        for _i, _step in enumerate(plan, 1):
            _q_raw = list(_step['joints'])
            _q_near = _nearest_in_limit(_q_raw)
            if _q_near != _q_raw:
                log('段%d 关节取同角等价表示：%s → %s'
                    % (_i, ['%.2f' % v for v in _q_raw], ['%.2f' % v for v in _q_near]))
                _step['joints'] = _q_near[:]          # 执行也用归一化值 ✓
            if not _real_limit_ok(_step['joints'], _lo, _hi):
                raise ValueError('段%d 目标关节超出实机限位：%s（规划期应已过滤，此为最后防线；已试 ±360 同角表示）'
                                 % (_i, ['%.2f' % v for v in _step['joints']]))
        for before, after in ((frame, robot.PoseFrame()), (tool, robot.PoseTool())):
            error = invH(before)*after
            if norm(error.Pos()) > 0.01 or pose_angle(error) > math.radians(0.01):
                raise RuntimeError('预检期间工具或参考坐标系改变，取消执行。')
        robot.setSpeed(ROBOT_SPEED)
        RDK.Command('Trace','Reset')
        RDK.Command('Trace','On')
        expected = start
        # v14k：停用长运动分瓣（split_moves 恒 False）。2026-10-12 实测日志坐实：假断连与跨度无关，
        # 60°/95°/169°/180° 的瓣与 20mm 途经点每条指令都在断，分瓣已不防任何东西，只剩每瓣一轮
        # 等待+重连停顿税；_single_move_settle 断连容忍（_wait_controller_static 20s 静止上限）
        # 罩得住单条长指令的收尾（20°/s 下 180°≈9s<20s）。分瓣机制与常量原样留档，遇真断连指纹
        # （未自然收尾/未到位）随时把本行改回 single_method is None and len(records) > 1 即可恢复。
        split_moves = False
        movl_direct = bool(real_movldirect_var.get()) if _movl_direct_ready() else False
        if movl_direct:
            # v15：原来的超长版本横幅已按用户要求删除，只留一行关键参数，便于判读
            log('直发开启 ｜ 段长≤%.0fmm ｜ 法兰容差 %.0fmm/%.1f° ｜ 等待≤%.0fs ｜ 禁直发名单=%s'
                % (MOVL_DIRECT_MAX_MM, MOVL_FLANGE_TOL_MM, MOVL_FLANGE_TOL_DEG,
                   MOVL_ARRIVE_WAIT_S, MOVL_DIRECT_BLOCK_POINTS))
        log('本次单条MovL动态认证放行点=%s' % [i for i,s in enumerate(plan,1) if s.get('direct_movl_certified')])
        _assert_continuous_dispatch(records, start, plan, movl_direct)
        for i, step in enumerate(plan, 1):
            for rewind in step['rewinds']:
                _require_joints(expected)
                _move_with_completion_check("MoveJ", rewind, split_moves)
                _require_joints(rewind)
                expected = rewind
            _require_joints(expected)
            waypoints = step.get('waypoints') or []
            if step['method'] == 'MoveL' and not waypoints:
                # 理论不可达：v13 起所有 MoveL 步都带细分途经点；不带则说明规划层契约被破坏
                raise RuntimeError(f"P{i}：MoveL 步缺少细分途经点，拒绝发送驱动 MOVL（已判死）。")
            seg_mm = seg_rot = None
            if movl_direct and step['method'] == 'MoveL' and waypoints:
                # 仅开关开启时才算（两次 FK 的 API 往返）；开关关/离线 verify 零开销
                _seg_rel = _trajectory_pose(step['joints']) * invH(_trajectory_pose(expected))
                seg_mm, seg_rot = norm(_seg_rel.Pos()), pose_angle(_seg_rel)
            direct_ready = (movl_direct and _direct_step_allowed(i, step)
                            and seg_mm is not None
                            and seg_mm <= MOVL_DIRECT_MAX_MM
                            and seg_rot <= math.radians(0.5))
            _send_q = step.get('direct_send_joints', step['joints'])
            if direct_ready and not step.get('direct_movl_certified'):
                # v14w：发送前数字净化——控制器 -30001 拒的是【参数形态】不是几何（LOG_VERSION
                # 处 11:38 拒收 / 15:55 接受两份实录）。净化只在零边界区微调发送关节；
                # 净化失败 ⇒ direct_ready=False ⇒ 落到 elif waypoints 走细分（安全回落）。
                _send_q, _purge_note = _movl_digit_safe_joints(step['joints'])
                if _send_q is None:
                    log('P%d：⛔ %s ⇒ 改走细分途经点路径。' % (i, _purge_note))
                    direct_ready = False
                elif _purge_note:
                    log('P%d：%s' % (i, _purge_note))
            if direct_ready:
                # v14p 法兰补偿MOVL：驱动 MOVL 无工具补偿、按法兰执行（v14l 11:30 实证停点法兰=
                # 命令TCP目标，差仅5.5mm）——将错就错：把本步构型的【法兰位姿】直接当笛卡尔目标
                # 发给控制器，法兰被精确送到位，物理工具尖端（182mm，v14w27 实测）随之落在认证
                # 直线上。姿态恒定段法兰线=TCP线平移常向量，扫掠包络与细分路径一致。
                # v14w36/37 演进：v14w36 只改传位姿（不切工具）⇒ MoveL(位姿) 按 TCP 空间
                # 校验，P8 法兰位姿被反推到 z=744 爆臂展 TargetReachError（11:18 实录）；
                # v14w37 = 位姿传递（动画=认证直线，根治关节弧假碰撞冻死）+ 发送窗口单位
                # 变换（校验/数字=法兰空间）；柜子实收参数与旧金标准逐位一致（0 偏差）。
                log(f"P{i}：v14w 法兰补偿MOVL：段长{seg_mm:.1f}mm（姿态变化{math.degrees(seg_rot):.2f}°），收起 {len(waypoints)} 个细分途经点，一指令直发（发法兰位姿=自算FK+单位变换窗口，发送关节已净化；v14w37）。")
                # v14r：require_joints=False——假断连分支的关节级 0.5° 校验让位给下方
                # 法兰级粗验收+MoveJ 微纠偏收口（终点仍回认证构型，护栏语义不降级）。
                # v14u：expect_target=段目标关节——目标锚定到位等待（上限 60s，每5s进度日志）。
                # v14w：净化只作用于发送关节；expect_target 仍是认证关节（到位判据不变）。
                # v14w37：位姿传递（动画=认证直线）+ flange_space 单位变换（校验/数字=法兰空间）。
                _send_pose = invH(robot.PoseFrame()) * robot.SolveFK(_send_q)
                # ★ 2026-11-03（可选，默认关）：先给控制器发 Tool(0)/User(0)，
                # 治 `[MovL#878] movL not set tool or user!!!` ⇒ 让 MovL 明确按 基座系+零工具(法兰) 执行。
                # 打开方式：把 MOVL_SEND_TOOL_USER 改成 True（建议先跑一条短段验证）。
                if MOVL_SEND_TOOL_USER:
                    if _try_set_tool_user():
                        log('  ✓ Tool(0)/User(0) 已下发，继续直发')
                    else:
                        raise ControllerMotionFault('Tool/User未确认，停止直发。')
                log('P%d：发送法兰目标=%s；认证关节=%s；TCP=%s' % (i, Pose_2_Fanuc(_send_pose), step['joints'], Pose_2_Fanuc(robot.PoseTool())))
                _single_move_settle('MoveL', _send_pose, require_joints=False,
                                    expect_target=step['joints'], flange_space=True)
                # ★★★ v15.7（2026-11-03）：直发结束后【先等真静止】再做后续（法兰验收/收口）。
                #   实录（v15.6, P8）：直发报"已完成"（假断连分支）→ 脚本立刻法兰验收(5.71mm ✓)
                #   → P8 尾部关节检查【通过】（读到的是过渡中姿态）→ P9 开头再读【已翻转】⇒ 差 20~38° ⇒ 停 ✗
                #   对比：P7 目标 [75.42,12.24,57.74,20.02] vs 停止实测 [78.10,36.86,19.48,33.66]
                #         ⇒ J2↑25 / J3↓38 / J4↑14 = 典型【肘部翻转 elbow flip】✗
                #   机理：MovL 只给位姿 ⇒ 控制器自行选 IK 分支（可能选翻转那组）✗
                #         + 直发"已完成"没等真静止 ⇒ 后续读到的是过渡值 ✗
                #   ⇒ 这里补一段【关节稳定等待】：连续 3 次采样（每次 0.3s）关节变化 <0.05° 才算真停，
                #     最多等 8 秒；等稳定后再做验收/收口，避免"读到过渡值"造成的假通过/假失败。
                _st = None
                _stable = False
                for _w in range(24):          # 24 × 0.3s ≈ 7.2s 上限
                    _cur = _live_joints()
                    if _st is not None and max(abs(a - b) for a, b in zip(_cur, _st)) < 0.05:
                        _stable = True
                        break
                    _st = _cur
                    time.sleep(0.3)
                if not _stable:
                    log('P%d：⚠️ 直发后 7 秒内关节仍未稳定（继续按现值验收，可能判死）' % i)
                else:
                    log('P%d：直发后关节已稳定 ✓（进入法兰验收/收口）' % i)
                # ★★★ v15.8（2026-11-03）：★ 安全网 —— 直发是【控制器自行选 IK 解】，
                #   规划期的自干涉硬禁区（|J4|>150 等）拦不到它 ✗
                #   ⇒ 直发落点若真落进禁区（J4 极端 / J4×J5 组合区），必须【立刻回认证构型】，
                #     绝不能把手臂留在危险姿态里继续跑下一段 ✓
                _post = _live_joints()
                if _real_interfere_combo(_post):
                    log('P%d：🚨 直发落点落入自干涉禁区！实测=%s（J4=%.2f J5=%.2f）⇒ 立即回认证构型'
                        % (i, ['%.2f' % v for v in _post], _post[3], _post[4]))
                    _single_move_settle('MoveJ', step['joints'])
                    _require_joints(step['joints'])
                    log('P%d：已回到认证构型 ✓' % i)
                elif abs(_post[3]) > REAL_INTERFERE_J4_MAX:
                    log('P%d：⚠️ 直发落点 J4=%.2f° 偏大（>%.0f° 组合区阈值，但未触禁区组合）——记录'
                        % (i, _post[3], REAL_INTERFERE_J4_MAX))
                try:
                    robot.setJoints(_post)   # 显示实测姿态，不用预期目标掩盖未到位。
                except Exception:
                    pass
                # v14q：MovL 落点法兰级粗验收（≤8mm/≤1°）+ MoveJ 微纠偏收口（关节级 0.5° 罩终点）。
                # v14p 首航停在 0.95° 关节残差（法兰 4.61mm/0.616°）被 0.5° 护栏拦停——那是控制器
                # MovL 固有落点残差（v14l 5.5mm 双样本背书），不是构型错误；但终点必须回到认证构型，
                # 故验收通过后用一条短 MoveJ（~1° 关节差）收口，走 _single_move_settle 全套护栏。
                _actual, _is_static = _wait_controller_static(samples=3, interval=0.2)
                _mm, _deg = _movl_flange_accept(_actual, step['joints'])
                if _mm > MOVL_FLANGE_TOL_MM or _deg > MOVL_FLANGE_TOL_DEG:
                    raise RuntimeError('v14u 法兰级粗验收未过：停点法兰残差%.2fmm/%.2f°（容差%.1fmm/%.1f°），实测关节%s，停止待判读。'
                                       % (_mm, _deg, MOVL_FLANGE_TOL_MM, MOVL_FLANGE_TOL_DEG,
                                          ['%.2f' % v for v in _actual]))
                _jm = max(abs(a - b) for a, b in zip(_actual, step['joints']))
                if _jm > MOVE_OFFSET_TOL:
                    log(f"P{i}：v14u MovL 直发落点法兰级验收通过（残差{_mm:.2f}mm/{_deg:.2f}°），关节残差{_jm:.2f}°——发 MoveJ 微纠偏收口。")
                    # ★★★ v15.4（2026-11-03）：收口 MoveJ 加重试 —— 治"P8 停下"：
                    #   实录 11:29:03 验收通过 → 发收口 MoveJ → 11:29:04 驱动报断连 → 11:29:06 才重连
                    #   ⇒ 那条收口 MoveJ 没走完 ⇒ 关节残差 2.68° 残留
                    #   ⇒ 下一段前的 _require_joints（容差 0.5°）判死 ⇒ 停在 P8 ✗
                    #   收口目标是【认证构型】（确定可达）⇒ 重发安全 ✓；最多 2 次，仍不到就抛原错。
                    _close_err = None
                    for _close_try in (1, 2):
                        try:
                            _single_move_settle('MoveJ', step['joints'])
                            _close_err = None
                            break
                        except Exception as _close_exc:  # noqa: BLE001
                            _close_err = _close_exc
                            if _close_try == 1:
                                log('P%d：收口 MoveJ 未完成（%s: %s）⇒ 重试一次（目标为认证构型，可达）'
                                    % (i, type(_close_exc).__name__, _close_exc))
                                time.sleep(0.5)
                    if _close_err is not None:
                        raise _close_err
                # ★★★ v15.5（2026-11-03）：直发+收口之后，再做【关节校正重试】—— 治 P8 停下的真因。
                #   实录（v15.4, 11:36:19~23）：
                #     P8 直发到位（关节残差 2.68°）→ 法兰验收通过 → 发收口 MoveJ
                #     → 驱动报断连 → 脚本打印「驱动断连但运动已自然完成到位」（★ 它认为完成 ✗）
                #     → 于是 _single_move_settle 没抛异常（断连分支 require_joints=False 不校验关节）
                #     → 紧接的 _require_joints 才发现不一致（实测 J2=36.86/J3=19.48，差很多）⇒ 抛错停 ✗
                #   ⇒ 所以 v15.4 的 try/except 重试【根本没触发】✗
                #   ⇒ 改为：_require_joints 失败时【再发一次定向 MoveJ】校正（目标=认证构型，确定可达）
                try:
                    _require_joints(step['joints'])
                except Exception:
                    log('P%d：直发+收口后关节仍与预检不一致 ⇒ 再发一次 MoveJ 校正（目标为认证构型，可达）' % i)
                    time.sleep(0.5)
                    _single_move_settle('MoveJ', step['joints'])
                    _require_joints(step['joints'])
                    log('P%d：校正 MoveJ 完成 ✓' % i)
            elif (movl_direct and not _direct_step_allowed(i, step) and seg_mm is not None
                    and seg_mm <= MOVL_DIRECT_MAX_MM and seg_rot <= math.radians(0.5)):
                # ★ v14v4：本点被【禁直发名单】拦下 —— 明确告知，便于判读日志
                log(f"P{i}：⛔ 本点在【禁直发名单】MOVL_DIRECT_BLOCK_POINTS={MOVL_DIRECT_BLOCK_POINTS} 里 ⇒ "
                    f"不走法兰补偿直发，改走【细分途经点路径】（v14n 实测 17/17 通过、零事故的路径）。")
                if not waypoints:
                    raise RuntimeError(f'P{i}：禁直发点缺少途经点，停止。')
                for way in waypoints:
                    _move_with_completion_check('MoveJ', way, False)
                    _require_joints(way)
                _require_joints(step['joints'])
            elif waypoints:
                log(f"P{i}：执行预检方案 {step['method']}→MoveJ 细分，{len(waypoints)} 个途经点，终点关节={step['joints']}")
                for k, way in enumerate(waypoints, 1):
                    _move_with_completion_check('MoveJ', way, False)
                    _require_joints(way)
                _require_joints(step['joints'])
            else:
                log(f"P{i}：执行预检方案 {step['method']}，关节={step['joints']}")
                _move_with_completion_check(step['method'], step['joints'], split_moves)
                _require_joints(step['joints'])
            expected = step['joints']
            completed += 1
        log(f'实机执行完成：{completed}/{len(plan)}点。')
    except Exception as exc:
        log(f'实机任务停止，已完成{completed}点：{type(exc).__name__}: {exc}')
        if movl_direct and ('断连' in str(exc) or '未到位' in str(exc) or '落点偏差' in str(exc) or '粗验收' in str(exc)):
            log('【v14u】法兰补偿MOVL执行段出断连/落点指纹（v14w24 无勾选框；细分途经点路径保留在计划中，可作回退依据）。')
        try:
            actual, velocity, mode = _controller_feedback()
            log('停止时控制器实际反馈：关节=%s，速度=%s，模式=%s；不自动重发运动。' % (actual, velocity, mode))
        except Exception as feedback_error:
            log('停止时也无法取得控制器反馈：%s' % feedback_error)
    finally:
        _real_running = False
        try:
            _keepalive_stop.set()
            _ka_thread.join(timeout=3)
        except Exception:
            pass


def _point_to_segment_distance(p, a, b):
    """3D点到线段距离，单位mm。"""
    ax, ay, az = a
    bx, by, bz = b
    px, py, pz = p
    ab = (bx-ax, by-ay, bz-az)
    ap = (px-ax, py-ay, pz-az)
    ab2 = ab[0]*ab[0] + ab[1]*ab[1] + ab[2]*ab[2]
    if ab2 < 1e-12:
        return math.sqrt((px-ax)**2 + (py-ay)**2 + (pz-az)**2)
    t = (ap[0]*ab[0] + ap[1]*ab[1] + ap[2]*ab[2]) / ab2
    t = max(0.0, min(1.0, t))
    q = (ax+t*ab[0], ay+t*ab[1], az+t*ab[2])
    return math.sqrt((px-q[0])**2 + (py-q[1])**2 + (pz-q[2])**2)


def _tcp_position_from_joints(q):
    """关节角 -> 当前参考坐标系下的TCP位置，与轨迹输入使用同一坐标系。"""
    f = pose_to_fanuc_values(invH(robot.PoseFrame()) * robot.SolveFK(q) * robot.PoseTool())
    return (float(f[0]), float(f[1]), float(f[2]))


def _check_movej_tcp_trajectory(start_q, target_q, start_tcp_vals, target_tcp_vals, log, samples=30, max_deviation_mm=None):
    """
    在真正执行MoveJ之前，用关节空间线性插补采样，计算TCP轨迹相对
    起点-终点TCP直线段的最大偏离距离。

    目的：MoveL失败时，不再无条件MoveJ；只有MoveJ造成的TCP空间绕行
    没有超过允许值，才允许用MoveJ兜底。
    """
    if max_deviation_mm is None:
        max_deviation_mm = MOVEJ_FALLBACK_MAX_DEVIATION_MM

    start_q = [float(v) for v in start_q[:6]]
    target_q = [float(v) for v in target_q[:6]]
    a = (float(start_tcp_vals[0]), float(start_tcp_vals[1]), float(start_tcp_vals[2]))
    b = (float(target_tcp_vals[0]), float(target_tcp_vals[1]), float(target_tcp_vals[2]))

    log("开始检查 MoveJ 兜底轨迹：%d 个采样点，允许最大TCP偏离 %.3f mm" % (samples + 1, max_deviation_mm))
    max_dev = -1.0
    max_info = None

    for k in range(samples + 1):
        t = float(k) / float(samples)
        q = [start_q[j] + (target_q[j] - start_q[j]) * t for j in range(6)]
        try:
            p = _tcp_position_from_joints(q)
        except Exception as e:
            log("  MoveJ轨迹检查失败：第 %d/%d 个采样点 FK失败：%s: %s" % (k+1, samples+1, type(e).__name__, e))
            return False

        dev = _point_to_segment_distance(p, a, b)
        if dev > max_dev:
            max_dev = dev
            max_info = (k, t, q, p)

        if dev > max_deviation_mm:
            log("✕ MoveJ兜底轨迹拒绝：第 %d/%d 个采样点偏离TCP直线 %.3f mm > %.3f mm" %
                (k+1, samples+1, dev, max_deviation_mm))
            log("  t=%.3f  TCP=(%.3f, %.3f, %.3f)" % (t, p[0], p[1], p[2]))
            log("  因此不会执行这个MoveJ兜底动作，避免出现不可接受的大绕圈。")
            return False

    if max_info is not None:
        k, t, q, p = max_info
        log("✓ MoveJ兜底轨迹检查通过")
        log("  最大TCP偏离直线：%.3f mm（采样 %d/%d，t=%.3f）" % (max_dev, k+1, samples+1, t))
        log("  最大偏离点TCP=(%.3f, %.3f, %.3f)" % (p[0], p[1], p[2]))
    return True


# ============================================================
# 执行连续运动（MoveL失败时先检查MoveJ轨迹）
# ============================================================
def _collision_details():
    pairs = RDK.CollisionPairs()
    return '；'.join(f'{a.Name()}[连杆{ia}] 与 {b.Name()}[连杆{ib}]'
                    for a, b, ia, ib in pairs) or '路径碰撞或关节不可行'


def _enable_obstacle_checks():
    if RDK.RunMode() != RUNMODE_SIMULATE:
        raise RuntimeError('障碍物预检仅允许在仿真模式执行。')
    # 每次进入预检都清空预检缓存：缓存生命周期 = 单次预检规划，
    # 障碍物/工作站状态的变化在下一次预检即时生效。
    _plan_cache.clear()
    for name in ('安装台_650x650x80mm', '地面_禁止穿越', '磨砂圆柱_R150_H50', '挡板_半封闭3面'):
        obstacle = RDK.Item(name, ITEM_TYPE_OBJECT)
        if not obstacle.Valid():
            raise RuntimeError(f'缺少障碍物模型：{name}，请加载包含台子和地面的工作站。')
        if name == '安装台_650x650x80mm':
            if RDK.setCollisionActivePair(COLLISION_OFF, robot, obstacle, 0, 0) != 1:
                raise RuntimeError('无法配置安装台与固定底座的接触关系。')
        for link in range(1, 7):
            if RDK.setCollisionActivePair(COLLISION_ON, robot, obstacle, link, 0) != 1:
                raise RuntimeError(f'无法启用{name}与连杆{link}的碰撞检查。')
        tool_items = list(RDK.ItemList(ITEM_TYPE_TOOL))
        _handle = RDK.Item('门把手_bs1')   # v14w12：网格替换后可能为 OBJECT 类型，按名并入
        if _handle.Valid() and all(_handle.item != t.item for t in tool_items):
            tool_items.append(_handle)
        for tool in tool_items:
            parent = tool.Parent()
            while parent.Valid() and parent.item != robot.item:
                parent = parent.Parent()
            if parent.Valid() and RDK.setCollisionActivePair(COLLISION_ON, tool, obstacle) != 1:
                raise RuntimeError(f'无法启用{name}与工具的碰撞检查。')
    RDK.setCollisionActive(COLLISION_ON)


def _check_single_joint_path(end):
    _enable_obstacle_checks()
    saved = robot.Joints().list()[:6]
    try:
        RDK.Command('Trace', 'Off')
        RDK.Render(False)
        if _movej_test_cached(saved, end, 1) != 0:
            raise ValueError('单点MoveJ路径被拒绝：' + _collision_details())
    finally:
        robot.setJoints(saved)
        RDK.Render(True)


def _trajectory_pose(q):
    return invH(robot.PoseFrame()) * robot.SolveFK(q) * robot.PoseTool()


def _reorient_next_pose(records, i, rec):
    """v14w33：i 为 1-based 点号。若下一点存在且为【同 TCP 位姿纯换姿】（xyz 全同、姿态不同），
    返回下一点的 TCP 位姿 Mat，否则 None。用于换姿对的分支前视。"""
    try:
        if i >= len(records):
            return None
        nxt = records[i]          # 0-based 列表：下一条记录
        if nxt['type'] != 'TCP' or nxt.get('singular', False):
            return None
        va = [float(v) for v in rec['values'][:6]]
        vb = [float(v) for v in nxt['values'][:6]]
        if all(abs(va[k] - vb[k]) < 1e-9 for k in range(3)) and any(abs(va[k] - vb[k]) > 1e-9 for k in range(3, 6)):
            return fanuc_values_to_pose(*vb)
    except Exception:
        return None
    return None


def _linear_path_endpoint(start, target):
    """带结果缓存：分支重试时同一（起点, 目标）不重复计算。"""
    key = ('linear', _cache_key_joints(start), _cache_key_pose(target))
    if key in _plan_cache:
        return _plan_cache[key]
    result = _linear_path_endpoint_uncached(start, target)
    _plan_cache[key] = result
    return result


def _linear_path_endpoint_uncached(start, target):
    # 粗筛：10mm 采样点是 1mm 采样点的子集，粗筛失败则 1mm 细查必然失败，
    # 可直接拒绝；粗筛通过后再跑原有 1mm 细查，通过/拒绝判定与只跑 1mm 完全一致。
    if RDK.RunMode() != RUNMODE_SIMULATE:
        raise RuntimeError('直线路径预检仅允许在仿真模式执行。')
    # v15.17: Lookahead may leave the model at the P10 wrist-spin posture.
    # RoboDK's numerical IK uses current model joints even with an explicit j1.
    # Reset the model seed before each independent path check.
    robot.setJoints(start)
    status = robot.MoveL_Test(start, target, minstep_mm=10)
    if status == 0:
        robot.setJoints(start)
        status = robot.MoveL_Test(start, target, minstep_mm=1)
    if status != 0:
        return None, f'MoveL原生路径检查未通过（{status}）：' + _collision_details()
    # 本机MoveL_Test返回成功后Joints()可能为全零；从插补矩阵读取实际终点。
    # 碰撞判定已由上方同路径 1mm MoveL_Test 完成，此处仅提取终点关节，
    # 关闭碰撞检查提速（实测约快两个数量级）；整段权威碰撞复核仍在
    # _verify_obstacle_plan（碰撞开、1mm）进行。
    program = RDK.AddProgram('_TCP仿真_路径预检', robot)
    try:
        program.setVisible(False)
        robot.setJoints(start)
        program.setPoseFrame(robot.PoseFrame())
        program.setPoseTool(robot.PoseTool())
        program.MoveJ(start)
        program.MoveL(target)
        message, matrix, status = program.InstructionListJoints(mm_step=1, deg_step=1, collision_check=COLLISION_OFF)
        if status < 0:
            return None, message
        end = matrix.tr().rows[-1][:6]
        error_pose = invH(target) * _trajectory_pose(end)
        if norm(error_pose.Pos()) > .01 or pose_angle(error_pose) > math.radians(.01):
            raise RuntimeError('路径预检返回的终点不匹配目标TCP。')
        return end, message
    finally:
        program.Delete()


def _linear_waypoints(start, target, step_mm=None):
    """v13：从一条 MoveL 指令采样细分途经关节点（按 IK 顺序，无分支翻转）。

    用 InstructionListJoints(mm_step=LINEAR_SUBSTEP_MM, collision_check=COLLISION_OFF) 采样：
    途经点与 MoveL 执行的是同一条几何直线，且 IK 连续选解（避免用全局 SolveIK 时
    途经点在多解间跳变）。碰撞已由 _linear_path_endpoint 的 MoveL_Test@1mm 权威判定，
    此处不再重复。返回含终点的关节点列表；空列表表示采样失败（调用方回退直达）。"""
    if step_mm is None:
        step_mm = LINEAR_SUBSTEP_MM
    key = ('waypoints', _cache_key_joints(start), _cache_key_pose(target), round(float(step_mm), 3))
    if key in _plan_cache:
        return [q[:] for q in _plan_cache[key]]
    program = RDK.AddProgram('_TCP仿真_细分采样', robot)
    saved = robot.Joints().list()[:6]
    try:
        program.setVisible(False)
        robot.setJoints(start)
        program.setPoseFrame(robot.PoseFrame())
        program.setPoseTool(robot.PoseTool())
        program.MoveJ(start)
        program.MoveL(target)
        message, matrix, status = program.InstructionListJoints(mm_step=step_mm, deg_step=1, collision_check=COLLISION_OFF)
        cols = matrix.tr().rows if matrix is not None else []
        if status < 0 or not cols:
            return []
        # 丢弃比步长更密的重复点（InstructionListJoints 在奇异附近会加密采样）
        picked = [list(map(float, cols[0][:6]))]
        for row in cols[1:]:
            q = list(map(float, row[:6]))
            if max(abs(a - b) for a, b in zip(q, picked[-1])) >= step_mm / 10.0:
                picked.append(q)
        # 去尾：InstructionListJoints 可能带比目标多一点的收尾点，以关节距离最近的为准
        end_q, _ = _linear_path_endpoint(start, target)
        if end_q is not None and picked and max(abs(a - b) for a, b in zip(end_q, picked[-1])) > 1.0:
            picked[-1] = list(map(float, end_q))
        _plan_cache[key] = [q[:] for q in picked]
        return [q[:] for q in picked]
    finally:
        program.Delete()
        robot.setJoints(saved)


def _obstacle_posture_key(q, reference=None):
    table = RDK.Item('安装台_650x650x80mm', ITEM_TYPE_OBJECT)
    height = 0.0
    if table.Valid():
        elbow = invH(table.PoseAbs()) * robot.PoseAbs() * robot.JointPoses(q)[3]
        height = elbow.Pos()[2]
    return (-round(height, 6), sum((v-r)**2 for v, r in zip(q, reference or [0]*6)), tuple(q))


def _obstacle_joint_target(start, values, max_deviation=None, log=None):
    """带结果缓存：同一（起点, 目标, 偏离上限）的兜底选解不重复搜索。"""
    key = ('obstacle', _cache_key_joints(start), tuple(round(float(v), 6) for v in values[:6]),
           round(float(max_deviation), 6) if max_deviation is not None else None)
    if key in _plan_cache:
        cached = _plan_cache[key]
        if isinstance(cached, ValueError):
            raise cached
        return cached
    try:
        result = _obstacle_joint_target_uncached(start, values, max_deviation, log)
    except ValueError as exc:
        _plan_cache[key] = exc
        raise
    _plan_cache[key] = result
    return result


def _obstacle_joint_target_uncached(start, values, max_deviation=None, log=None):
    # v14-P2P：不再用 seed 候选/肘高排序，直接取离当前关节最近的逆解做逐级检查；
    # 最近解过不了偏离/碰撞时仍会在这里报错（单点 MoveJ 兜底路径保持可用）。
    lower, upper, _ = robot.JointLimits()
    candidates = [_nearest_ik_from_current(start, fanuc_to_pose(*values))]
    saved = robot.Joints().list()[:6]
    try:
        # 少量FK采样仅用于排序；不能替代后面的偏离复核与精细碰撞检查。
        a = _tcp_position_from_joints(start)
        table = RDK.Item('安装台_650x650x80mm', ITEM_TYPE_OBJECT)
        base_to_table = invH(table.PoseAbs()) * robot.PoseAbs()
        ranked = []
        for end in candidates:
            deviation, height = 0.0, float('inf')
            for k in range(11):
                q = [x + (y-x)*k/10 for x, y in zip(start, end)]
                deviation = max(deviation, _point_to_segment_distance(
                    _tcp_position_from_joints(q), a, values[:3]))
                height = min(height, (base_to_table * robot.JointPoses(q)[3]).Pos()[2])
            if max_deviation is not None and deviation > max_deviation:
                continue
            # 20mm一档，避免为很小的偏离差反复搜索；同档优先抬高肘部。
            ranked.append(((int(deviation/20), -height,
                            sum(abs(y-x) for x, y in zip(start, end))), end))
        checked = 0
        for _, end in sorted(ranked, key=lambda entry: entry[0]):
            if max_deviation is not None and not _check_movej_tcp_trajectory(
                    start, end, pose_to_fanuc_values(_trajectory_pose(start)), values,
                    lambda msg: None, samples=100, max_deviation_mm=max_deviation):
                continue
            checked += 1
            if _movej_test_cached(start, end, .25) == 0:
                if log is not None:
                    log(f'MoveJ快速筛选：{len(candidates)}个候选，{len(ranked)}个通过粗筛，精查{checked}条后找到合格路径。')
                return end
        raise ValueError('所有候选关节路径均碰撞、超出偏离限制或没有有效逆解。')
    finally:
        robot.setJoints(saved)


def _verify_obstacle_plan(start, plan):
    program = RDK.AddProgram('_TCP仿真_整段碰撞复核', robot)
    saved = robot.Joints().list()[:6]
    try:
        program.setVisible(False)
        program.setPoseFrame(robot.PoseFrame())
        program.setPoseTool(robot.PoseTool())
        program.MoveJ(start)
        for step in plan:
            for q in step['rewinds']:
                program.MoveJ(q)
            if step['method'] == 'MoveL' and not step.get('waypoints'):
                # v13 防呆：MoveL 步必须带细分途经点，否则规划层契约被破坏
                raise ValueError('整段碰撞复核：MoveL 步缺少细分途经点，拒绝。')
            getattr(program, step['method'])(step['joints'])
        message, matrix, status = program.InstructionListJoints(
            mm_step=1, deg_step=1, collision_check=COLLISION_ON)
        if status < 0 or 'collision' in message.lower():
            raise ValueError('整段碰撞复核未通过：' + message)
    finally:
        program.Delete()
        robot.setJoints(saved)


# Continuous TCP paths always recover calibrated-body IK branches and re-certify
# their actual command paths. Record hashes bind receipts, never enable policy.
CALIBRATED_IK_SEEDS = [[163.62039271007563, 64.01735255223417, -67.25050650734438, 93.2331539551102, -90.00000000000001, -106.37960728992437], [-72.40715810734315, -20.66480267505412, -103.89758096136477, 124.56238363641887, 72.40715810734312, 0.0], [-58.553344176794326, -22.475689666466394, -101.12528805253322, 123.60097771899962, 58.55334417679429, -1.0294949594003553e-14], [-58.553344176794326, -22.475689666466394, -101.12528805253322, 123.60097771899962, 58.55334417679429, 180.0], [-87.40476475829131, -22.47568966646641, -101.12528805253322, 123.60097771899962, 87.40476475829125, 180.0], [-64.66430037296594, -3.2481937678895747, -126.71804809984242, 129.96624186773198, 64.66430037296595, 180.0], [-75.41679324948196, -12.462263518678185, -56.77419042193441, -20.76354605938741, 90.0, 194.58320675051806], [-78.10373775148642, -37.83824919659381, -16.865010237740023, -35.296740565666134, 90.0, 191.89626224851355], [-88.23587605840977, -43.75520866199254, -5.060724146438354, -41.184067191569056, 90.0, 181.7641239415902], [-88.23587605840977, -43.75520866199254, -5.060724146438354, -41.184067191569056, 90.0, 1.7641239415902135], [-68.33462268250656, -43.75520866199333, -5.060724146436616, -41.184067191570016, 89.99999999999999, 21.665377317493437], [61.81374704354286, 48.51918849734889, 55.392423259627606, -103.91161175697648, 28.186252956457167, 180.0], [62.25330564679723, 54.06615976151417, 44.56648765802543, -98.6326474195396, 27.746694353202802, 180.0], [61.81374704354286, 48.51918849734889, 55.392423259627606, -103.91161175697648, 28.186252956457167, 90.0], [62.253305646797244, 54.06615976151415, 44.56648765802541, -98.63264741953954, 27.746694353202788, 89.99999999999999], [61.81374704354286, 48.51918849734889, 55.392423259627606, -103.91161175697648, 28.18625295645714, -90.00000000000001], [62.25330564679723, 54.0661597615141, 44.56648765802556, -98.63264741953965, 27.746694353202773, -90.00000000000004], [62.57433490659918, 47.78974891048301, 57.14855554302247, -103.76676871515006, 27.416346223420135, -60.70732349501101], [62.98154845233014, 53.155168153175346, 46.7150047327387, -98.68233310181975, 27.009218983764953, -60.72565665513798], [62.57582549469282, 48.080389017894106, 56.23528280269005, -104.31567182058413, 27.424174505307207, -180.0], [62.71034615480792, 51.83128832842894, 49.315963732196764, -99.89133677590429, 25.437207443150072, -301.4668568689523], [60.218467190004304, 39.42913510297621, 54.58098026787218, -92.8583848548389, 27.92853761288419, -301.35028218541504], [-13.591622773947876, 18.9460252211274, 48.02925373146127, 23.02472104741136, -90.0, -193.59162277394785]]
_continuous_profile_active = False


def _records_fingerprint(records):
    import hashlib
    canonical = [dict(type=r['type'], values=[0.0 if abs(float(v)) < 1e-12 else float(v)
                 for v in r['values']], singular=bool(r.get('singular', False)),
                 spin360=bool(r.get('spin360', False)), j6_delta=int(r.get('j6_delta', 0)))
                 for r in records]
    return hashlib.sha256(json.dumps(canonical, sort_keys=True,
        separators=(',', ':')).encode('utf-8')).hexdigest()


def _continuous_records(records):
    return len(records) > 1 and any(r.get('type') == 'TCP' for r in records)


def _assert_continuous_dispatch(records, initial, plan, direct_enabled):
    if not _continuous_records(records):
        return
    fingerprint = _records_fingerprint(records)
    previous = initial
    for number, step in enumerate(plan, 1):
        if step.get('waypoints'):
            certificate = step.get('direct_certificate') or {}
            if (step['method'] != 'MoveL' or not step.get('direct_movl_certified')
                    or certificate.get('records_sha256') != fingerprint
                    or certificate.get('start_joints') != list(previous)
                    or certificate.get('end_joints') != step['joints']
                    or certificate.get('send_joints') != step.get('direct_send_joints')):
                raise RuntimeError(f'P{number}缺少与当前数据及构型一致的连续直线认证，禁止退回逐点停走。')
            if not direct_enabled:
                raise RuntimeError('连续TCP轨迹需要单条MovL模式，禁止退回细分停走。')
        previous = step['joints']


def _controller_body_matches():
    expected = Fanuc_2_Pose([1.119989104069524, -245.1846134160959,
        1047.9330384567963, -89.7671431696512, -0.00006721956284782927,
        179.8638590144166])
    err = invH(expected) * robot.SolveFK([0.0] * 6)
    return norm(err.Pos()) < .001 and pose_angle(err) < math.radians(.001)


def _profile_ik_all(flange):
    native = robot.SolveIK_All(flange)
    if not _continuous_profile_active:
        return native
    key = ('profile_ik', _cache_key_pose(flange))
    if key in _plan_cache:
        return _plan_cache[key]
    raw = [list(q[:6]) for q in native]
    for seed in CALIBRATED_IK_SEEDS:
        q = robot.SolveIK(flange, seed).list()
        if len(q) >= 6:
            raw.append(q[:6])
    valid = []
    for q in raw:
        if len(q) != 6:
            continue
        q = [(float(v) + 180.0) % 360.0 - 180.0 for v in q]
        err = invH(flange) * robot.SolveFK(q)
        if norm(err.Pos()) > .001 or pose_angle(err) > math.radians(.001):
            continue
        if not any(max(abs(x-y) for x, y in zip(q, old)) < .001 for old in valid):
            valid.append(q)
    result = Mat(valid).tr() if valid else Mat(6, 0)
    _plan_cache[key] = result
    return result


def _direct_step_allowed(number, step):
    return number not in MOVL_DIRECT_BLOCK_POINTS or bool(step.get('direct_movl_certified'))


def _certify_continuous_direct(records, initial, plan, log):
    if not _continuous_profile_active:
        return
    if RDK.RunMode() != RUNMODE_SIMULATE or not _controller_body_matches():
        raise RuntimeError('本体或模式与连续TCP单条MovL验证条件不一致。')
    pose, link, frame, saved = robot.PoseTool(), robot.getLink(ITEM_TYPE_TOOL), robot.PoseFrame(), robot.Joints().list()[:6]
    lower, upper, _ = robot.JointLimits()
    try:
        for number, step in enumerate(plan, 1):
            if step['method'] != 'MoveL':
                continue
            if step['method'] != 'MoveL' or not step.get('waypoints'):
                raise ValueError(f'P{number}未形成连续直线，禁止以MoveJ代替本次工艺段。')
            start = initial if number == 1 else plan[number-2]['joints']
            relative = _trajectory_pose(step['joints']) * invH(_trajectory_pose(start))
            if norm(relative.Pos()) > MOVL_DIRECT_MAX_MM or pose_angle(relative) > math.radians(.5):
                raise ValueError(f'P{number}将退回{len(step["waypoints"])}段停走，换入口分支重试。')
            send_q, note = _movl_digit_safe_joints(step['joints'])
            if send_q is None:
                raise ValueError(f'P{number}发送位姿净化失败。')
            target = invH(frame) * robot.SolveFK(send_q)
            flange_tool = _named_tool(FLANGE_TOOL_NAME, eye(4))
            robot.setPoseTool(flange_tool)
            robot.setJoints(start)
            if robot.MoveL_Test(start, target, minstep_mm=.5) != 0:
                raise ValueError(f'P{number}净化后的法兰直线碰撞或不可达。')
            program = RDK.AddProgram('_轨迹16_单条MovL复核', robot)
            try:
                program.setVisible(False)
                program.setPoseTool(eye(4))
                program.setPoseFrame(frame)
                program.MoveJ(start)
                program.MoveL(send_q)
                robot.setJoints(start)
                message, matrix, status = program.InstructionListJoints(
                    mm_step=.5, deg_step=.2, collision_check=COLLISION_ON)
                samples = matrix.tr().rows
                if status < 0 or 'collision' in message.lower() or not samples:
                    raise ValueError(f'P{number}法兰整段复核失败：{message}')
                for row in samples:
                    q = row[:6]
                    if (int(row[6]) != 0 or not _real_limit_ok(q, lower.list(), upper.list())
                            or _real_interfere_combo(q)):
                        raise ValueError(f'P{number}法兰路径存在错误、限位或自干涉。')
                if max(abs(a-b) for a, b in zip(samples[-1][:6], send_q)) > .05:
                    raise ValueError(f'P{number}法兰直线落点分支与认证关节不一致。')
                err = invH(robot.SolveFK(send_q)) * robot.SolveFK(samples[-1][:6])
                if norm(err.Pos()) > .01 or pose_angle(err) > math.radians(.01):
                    raise ValueError(f'P{number}法兰路径终点不匹配。')
                step['direct_movl_certified'] = True
                step['direct_send_joints'] = list(send_q)
                step['direct_certificate'] = dict(records_sha256=_records_fingerprint(records),
                    start_joints=list(start), end_joints=list(step['joints']), send_joints=list(send_q),
                    samples=len(samples), flange_target=Pose_2_Fanuc(target), digit_note=note)
                log(f'P{number}：单条法兰MovL复核通过（0.5mm采样、碰撞/实机限位/落点分支）；本次免除细分。')
            finally:
                program.Delete()
                _restore_tool(pose, link)
    finally:
        _restore_tool(pose, link)
        robot.setPoseFrame(frame)
        robot.setJoints(saved)


def _ik_branch_candidates(target_pose, reference):
    """v14c：某个 TCP 位姿的全部限位内 IK 分支（含 J6 圈数取近表示），
    与 _nearest_ik_from_current 同款筛选规则。"""
    solutions = _profile_ik_all(_tcp_target_to_flange(target_pose))
    lower, upper, _ = robot.JointLimits()
    lower, upper = lower.list(), upper.list()
    candidates = []
    for solution in solutions:
        q = [((float(v) + 180.0) % 360.0) - 180.0 for v in solution[:6]]
        if len(q) != 6:
            continue
        for turns6 in (0, -1, 1):
            candidate = q[:]
            candidate[5] += 360.0 * turns6
            if _real_limit_ok(candidate, lower, upper):
                if not any(max(abs(a-b) for a, b in zip(candidate, old)) < 1e-6 for old in candidates):
                    candidates.append(candidate)
    for q in candidates[:]:
        nearest = [min((v + 360*k for k in range(math.ceil((lower[j]-v)/360),
                       math.floor((upper[j]-v)/360)+1)), key=lambda a: abs(a-reference[j]))
                   for j, v in enumerate(q)]
        # v14w22：取近表示必须复核实机限位（此前漏检 ⇒ J1=193.59 混入实发被 -40001 拒）
        if not _real_limit_ok(nearest, lower, upper):
            continue
        if not any(max(abs(a-b) for a, b in zip(nearest, old)) < 1e-6 for old in candidates):
            candidates.append(nearest)
    return candidates


def _nearest_ik_from_current_lookahead(current_q, target_pose, lookahead_ok):
    """v14i：同 _nearest_ik_from_current，但要求选出的解能满足前视条件 lookahead_ok(cand)->bool；
    没有满足者时退回最近解（死路由后续救援链/种子重试兜底）。"""
    candidates = _ik_branch_candidates(target_pose, current_q)
    if not candidates:
        raise ValueError('没有限位内的逆解。')
    ranked = sorted(candidates, key=lambda q: sum((q[j]-current_q[j])**2 for j in range(6)))
    for cand in ranked:
        if lookahead_ok(cand):
            return cand[:]
    return ranked[0][:]


def _nearest_ik_from_current(current_q, target_pose):
    """v14-P2P：从全部逆解中选离当前关节角最近的解（含 J6 圈数取近）。

    与 test.py 的肘高排序不同：以【关节空间离当前构型最近】为准，相邻点之间不会突变构型。
    没有限位内解时抛 ValueError。"""
    solutions = _profile_ik_all(_tcp_target_to_flange(target_pose))
    lower, upper, _ = robot.JointLimits()
    lower, upper = lower.list(), upper.list()
    candidates = []
    for solution in solutions:
        q = [((float(v) + 180.0) % 360.0) - 180.0 for v in solution[:6]]
        if len(q) != 6:
            continue
        for turns6 in (0, -1, 1):
            candidate = q[:]
            candidate[5] += 360.0 * turns6
            if _real_limit_ok(candidate, lower, upper):
                if not any(max(abs(a-b) for a, b in zip(candidate, old)) < 1e-6 for old in candidates):
                    candidates.append(candidate)
    # 同一姿态再补一圈数取近的表示，避免强制归零导致大绕行。
    for q in candidates[:]:
        nearest = [min((v + 360*k for k in range(math.ceil((lower[j]-v)/360),
                       math.floor((upper[j]-v)/360)+1)), key=lambda a: abs(a-current_q[j]))
                   for j, v in enumerate(q)]
        # v14w22：取近表示必须复核实机限位（此前漏检 ⇒ J1=193.59 混入实发被 -40001 拒）
        if not _real_limit_ok(nearest, lower, upper):
            continue
        if not any(max(abs(a-b) for a, b in zip(nearest, old)) < 1e-6 for old in candidates):
            candidates.append(nearest)
    if not candidates:
        raise ValueError('没有限位内的逆解。')
    return min(candidates, key=lambda q: sum((q[j]-current_q[j])**2 for j in range(6)))[:]


def _checked_j6_rewinds(q, lower, upper, max_deviation):
    """返回可实际执行的整圈回绕列表（带缓存）；TCP空间偏离和碰撞都必须通过检查。"""
    key = ('rewinds', _cache_key_joints(q), tuple(round(float(v), 6) for v in lower[:6]),
           tuple(round(float(v), 6) for v in upper[:6]), round(float(max_deviation), 6))
    if key in _plan_cache:
        return [r[:] for r in _plan_cache[key]]
    results = []
    tcp = pose_to_fanuc_values(_trajectory_pose(q))
    for delta in (-360.0, 360.0):
        end = q[:]
        end[5] += delta
        if not lower[5] <= end[5] <= upper[5]:
            continue
        if not _check_movej_tcp_trajectory(q, end, tcp, tcp, lambda msg: None,
                                          samples=360, max_deviation_mm=max_deviation):
            continue
        if _movej_test_cached(q, end, 1) == 0:
            results.append(end)
    _plan_cache[key] = results
    return [r[:] for r in results]


def _plan_continuous_trajectory(records, max_deviation, log):
    """v14c：首点全分支种子枚举 + 整段重试。

    贪心最近解在换向步（如轨迹7 P6 的原地转 90°→180°）会把 wrist 构型选到贴圆柱，
    后续任何分支都碰；TCP仿真宏靠首点种子枚举+整段重试避开这类死路。v14c 移植该机制：
    种子按肘高排序优先，贪心只负责段内选解；某段死路（含 MoveL 兑底都失败）
    则整段换种子重试，全部种子失败才报错。"""
    global _preferred_seed, _continuous_profile_active
    _continuous_profile_active = False
    if _continuous_records(records):
        if not _controller_body_matches():
            raise RuntimeError('连续TCP轨迹策略要求控制器对齐本体；当前本体参数不符。')
        if not _same_tool_pose(robot.PoseTool(), Fanuc_2_Pose(list(CANONICAL_TOOL))):
            raise RuntimeError('连续TCP轨迹策略要求130mm TCP。')
        if norm(robot.PoseFrame().Pos()) > .01 or pose_angle(robot.PoseFrame()) > math.radians(.01):
            raise RuntimeError('连续TCP轨迹策略要求机器人基座参考系。')
        _continuous_profile_active = True
        log('v15.22：启用校准本体分支搜索及防停走检查；不依赖旧坐标指纹，全部直线按当前数据重新认证。')
    _enable_obstacle_checks()
    if not math.isfinite(max_deviation) or max_deviation < 0:
        raise ValueError('MoveJ允许偏离必须是非负有限数。')
    for i, rec in enumerate(records):
        vals = rec['values']
        if rec['type'] not in ('TCP', 'JOINT') or len(vals) != 6 or not all(math.isfinite(v) for v in vals):
            raise ValueError(f'P{i+1}：点类型或六维数值无效。')
        if rec.get('singular', False):
            # v14a：恢复 v13 同款奇异点规则校验（P2P 规划层支持奇异点步）
            if rec['type'] != 'TCP' or i == 0 or records[i-1]['type'] != 'TCP' or records[i-1].get('singular', False):
                raise ValueError(f'P{i+1}：特异点必须紧跟普通TCP点。')
            if rec.get('spin360', False):
                if rec.get('j6_delta', 360) not in (-360, 360):
                    raise ValueError(f'P{i+1}：J6自转方向必须为+360或-360。')
                if max(abs(a - b) for a, b in zip(rec['values'], records[i-1]['values'])) > 1e-3:
                    raise ValueError(f'P{i+1}：J6自转360°特异点的六维数值必须与前一个TCP点完全相同。')
            elif rec.get('j6_delta', 180) not in (-180, 180):
                raise ValueError(f'P{i+1}：J6方向必须为+180或-180。')
    saved = robot.Joints().list()[:6]
    lower, upper, _ = robot.JointLimits()
    lower, upper = lower.list(), upper.list()
    # 先检查点本身可达，避免后面的不可达点触发整段分支重复搜索。
    unreachable = []
    for i, rec in enumerate(records, 1):
        if rec['type'] == 'TCP' and not rec.get('singular', False):
            target = fanuc_values_to_pose(*rec['values'])
            if _profile_ik_all(_tcp_target_to_flange(target)).size(1) == 0:
                unreachable.append(f'P{i}：没有逆解；' + _flange_target_description(target))
    if unreachable:
        raise ValueError('目标点不可达，尚未搜索连接路径：' + '；'.join(unreachable))
    if _movej_test_cached(saved, saved, 1) != 0:
        raise ValueError('起始姿态已碰撞，不能自动规划脱离：' + _collision_details())
    try:
        RDK.Render(False)
        # v14c：首点全分支种子枚举（肘高优先），某种子整段死路时换构型重试。
        first_tcp = next((r for r in records if r['type'] == 'TCP' and not r.get('singular', False)), None)
        if first_tcp is not None:
            seeds = _ik_branch_candidates(fanuc_values_to_pose(*first_tcp['values']), saved)
            seeds.sort(key=lambda s: _obstacle_posture_key(s, saved))
            if _continuous_profile_active:
                # Recover the previously successful entry branch on this calibrated body.
                # These are IK seeds, never executable joint targets.
                entry = robot.SolveIK(_tcp_target_to_flange(
                    fanuc_values_to_pose(*first_tcp['values'])), CALIBRATED_IK_SEEDS[0]).list()
                if len(entry) == 6:
                    seeds.sort(key=lambda s: sum((a-b)**2 for a,b in zip(s, entry)))
                log('v15.22：优先历史成功入口分支；任何细分停走退化均重新选解或停止预检。')
        else:
            seeds = [None]
        seed_context = repr((records, saved, robot.PoseFrame().rows, robot.PoseTool().rows, max_deviation))
        if _preferred_seed is not None and _preferred_seed[0] == seed_context:
            preferred = _preferred_seed[1]
            seeds.sort(key=lambda s: 0 if s == preferred else 1)
            log('优先尝试上次通过的首点构型；本次所有碰撞与整段检查仍重新执行。')
        last_seed_error = None
        for seed_rank, seed in enumerate(_lazy_valid_seeds(seeds, saved), 1):
            if len(seeds) > 1:
                log(f'—— 尝试首点分支种子 {seed_rank}/{len(seeds)}：' +
                    ('%s' % [round(v, 1) for v in seed] if seed else '无种子(关节轨迹)'))
            q = saved[:]
            plan = []
            try:
                seed_used = seed is None
                for i, rec in enumerate(records, 1):
                    rewinds = []
                    delta = None
                    method, fallback, waypoints = 'MoveJ', False, []
                    lookahead_ok = None  # v14j：循环顶初始化（首个TCP点走种子路径时前视绑定也可安全引用）
                    if rec['type'] == 'JOINT':
                        end = [float(v) for v in rec['values'][:6]]
                        note = '录入关节直达'
                    elif rec.get('singular', False):
                        # v14a：奇异点步——只转 J6（±180 换向 / ±360 自转）。
                        # ±180：从当前解纯转 J6，由下方 FK 校验把关；超限时先试反方向（终点位姿不变）再试整圈回绕。
                        target = fanuc_values_to_pose(*rec['values'])
                        delta = rec.get('j6_delta', 180)

                        def _fk_matches(candidate):
                            error_pose = invH(target) * _trajectory_pose(candidate)
                            return norm(error_pose.Pos()) <= 1e-3 and pose_angle(error_pose) <= math.radians(.01)

                        end = q[:]
                        end[5] += delta
                        if not lower[5] <= end[5] <= upper[5]:
                            alt = q[:]
                            alt[5] -= delta
                            if lower[5] <= alt[5] <= upper[5]:
                                log(f'P{i}：J6 {delta:+d}°超限，改用反方向 {-delta:+d}°（终点位姿不变）。')
                                end, delta = alt, -delta
                            if not lower[5] <= end[5] <= upper[5]:
                                for rewound in _checked_j6_rewinds(q, lower, upper, max_deviation):
                                    if lower[5] <= rewound[5] + delta <= upper[5]:
                                        rewinds.append(rewound[:])
                                        q = rewound
                                        end = q[:]
                                        end[5] += delta
                                        break
                                else:
                                    raise ValueError(f'P{i}：J6 {delta:+d}°超限：反方向与整圈回绕均不可行。')
                        if not _fk_matches(end):
                            raise ValueError(f'P{i}：仅旋转J6无法到达所标注TCP，请检查特异点标记/工具。')
                        # v14d：换向步碰撞时，先试反方向（终点位姿不变），再试整圈回绕——
                        # TCP仿真靠方向枚举能避开这类碰撞，P2P 此前只在超限时才换向。
                        # v14j：反方向终点=当前解−delta（旧代码误算 q−2δ，朝向未翻转、FK 必不匹配，
                        # 15/15 种子全死于此——probe_p14_lookahead.py 坐实）。
                        if _movej_test_cached(q, end, 1) != 0:
                            alt = q[:]
                            alt[5] -= delta
                            flipped = False
                            if lower[5] <= alt[5] <= upper[5] and _fk_matches(alt) and _movej_test_cached(q, alt, 1) == 0:
                                log(f'P{i}：J6 {delta:+d}°扫过障碍，改用反方向 {-delta:+d}°（终点位姿不变）。')
                                end, delta, flipped = alt, -delta, True
                            if not flipped:
                                for rewound in _checked_j6_rewinds(q, lower, upper, max_deviation):
                                    cand = rewound[:]
                                    cand[5] += delta
                                    if lower[5] <= cand[5] <= upper[5] and _fk_matches(cand) and _movej_test_cached(q, cand, 1) == 0:
                                        log(f'P{i}：J6 {delta:+d}°两方向均碰，先整圈回绕再换向。')
                                        rewinds.append(rewound[:])
                                        q, end, flipped = rewound, cand, True
                                        break
                            if not flipped:
                                # v14f：两方向都碰——先切到同位姿的其他 IK 分支（碰撞预检过），
                                # 从那里再换向；途经的构型跳记入 rewinds 由执行层逐跳执行。
                                # v14j：枚举基准改为当前（未翻转）位姿——旧代码误用翻转后 target，
                                # 候选再 ±180 回到未翻转位姿，FK 对 target 永不匹配，结构性必死。
                                for cand in sorted(_ik_branch_candidates(_trajectory_pose(q), q),
                                                   key=lambda c: sum((c[j]-q[j])**2 for j in range(6))):
                                    for sgn in (delta, -delta):
                                        after = cand[:]
                                        after[5] += sgn
                                        if not (lower[5] <= after[5] <= upper[5] and _fk_matches(after)):
                                            continue
                                        if _movej_test_cached(q, cand, 1) == 0 and _movej_test_cached(cand, after, 1) == 0:
                                            log(f'P{i}：J6 ±180°两方向均碰，先切IK分支再换向（rewinds 跳转）。')
                                            rewinds.append(cand[:])
                                            q, end, delta, flipped = cand, after, sgn, True
                                            break
                                    if flipped:
                                        break
                            if not flipped:
                                # v14g：同位姿先 MoveL 到场再换向——MoveL 连续选解给出的构型
                                # 正是 TCP仿真 实测可换向的构型（贪心最近解构型两方向都扫障碍）。
                                lin_end, lin_detail = _linear_path_endpoint(q, target)
                                if lin_end is not None:
                                    pre_waypoints = _linear_waypoints(q, target)
                                    if pre_waypoints:
                                        for sgn in (delta, -delta):
                                            after = lin_end[:]
                                            after[5] += sgn
                                            if not (lower[5] <= after[5] <= upper[5] and _fk_matches(after)):
                                                continue
                                            if _movej_test_cached(lin_end, after, 1) == 0:
                                                log(f'P{i}：J6 两方向均碰，先 MoveL 到场（连续选解构型）再{sgn:+d}°换向。')
                                                plan.append(dict(method='MoveL', joints=lin_end[:], special=False,
                                                                 fallback=False, rewinds=[], j6_delta=None,
                                                                 waypoints=pre_waypoints, p2p_note='换向前MoveL到场'))
                                                q, end, delta, flipped = lin_end[:], after, sgn, True
                                                break
                            if not flipped:
                                raise ValueError(f'P{i}：J6 ±180°换向两方向均碰撞（含回绕/分支/MoveL到场尝试），该构型不可行。')
                        note = ('J6自转%+d°' % delta) if rec.get('spin360', False) else ('J6换向%+d°' % delta)
                    else:
                        target = fanuc_values_to_pose(*rec['values'])
                        # v14h：与前一点同位姿（停顿点，如轨迹7 P7）——不重新选解，
                        # 保持当前构型不动，只往计划里记一个停顿点。
                        if max(abs(_trajectory_pose(q).Pos()[j] - target.Pos()[j]) for j in range(3)) < 1e-3 and \
                           pose_angle(invH(target) * _trajectory_pose(q)) < math.radians(.01):
                            plan.append(dict(method='MoveJ', joints=q[:], special=False, fallback=False,
                                             rewinds=[], j6_delta=None, waypoints=[], p2p_note='同位姿停顿'))
                            continue
                        if not seed_used:
                            end = seed[:]  # v14c：首个TCP点直接采用种子分支（离起点可达性已在种子筛选时验证）
                            seed_used = True
                        else:
                            # v14i：前视——下一个执行点是 ±180 换向时，本点选解必须能完成那次换向
                            #（两方向任一可通行），否则贪心构型会把换向逼成死路。
                            nxt = records[i] if i < len(records) else None
                            lookahead_ok = None
                            if nxt is not None and nxt.get('singular', False) and not nxt.get('spin360', False):
                                nxt_values = nxt['values']
                                def lookahead_ok(cand, _vals=nxt_values, _lower=lower, _upper=upper):
                                    nxt_target = fanuc_values_to_pose(*_vals)
                                    for sgn in (180, -180):
                                        after = cand[:]
                                        after[5] += sgn
                                        if not (_lower[5] <= after[5] <= _upper[5]):
                                            continue
                                        err = invH(nxt_target) * _trajectory_pose(after)
                                        if norm(err.Pos()) > 1e-3 or pose_angle(err) > math.radians(.01):
                                            continue
                                        if _movej_test_cached(cand, after, 1) == 0:
                                            return True
                                    return False
                                log(f'P{i}：前视模式（P{i+1}为±180换向，选解需兼顾换向可行性）。')
                            end = (_nearest_ik_from_current_lookahead(q, target, lookahead_ok)
                                   if lookahead_ok else _nearest_ik_from_current(q, target))
                        note = 'TCP最近解直达'
                        forced_lin = False
                        # v14w24：短直线工作段强制 MoveL——P2→P3 这类 ≤210mm/姿态恒定 的
                        # 贴面平移，工艺不允许 MoveJ 关节弧绕行，直走直线（判据与直发门禁同款）。
                        # 前视夜（下一点±180换向）：直线末端同样具备换向资格才强制，否则回落
                        # MoveJ 前视绑定（保住换向可行性纪律）。
                        _rel = _trajectory_pose(q) * invH(target)
                        _seg_mm_f = norm(_rel.Pos())
                        _force_ok = _seg_mm_f <= MOVL_DIRECT_MAX_MM and pose_angle(_rel) <= math.radians(0.5)
                        # v14w33c：回撤段（TCP y 朝基座 >10mm）且下一点是同位姿换姿 ⇒ 让位 MoveJ
                        # 分支前视（强制 MoveL 的端点分支由直线 IK 连续性锁死，会对下一点无路：
                        # P5→P6→P7 实录 P7 被迫 49 跳细分）。工艺贴面滑移（Δy≈0）不受影响。
                        if _force_ok and i >= 2 and _reorient_next_pose(records, i, rec) is not None:
                            try:
                                _y_prev = float(records[i - 2]['values'][1])
                                if float(rec['values'][1]) - _y_prev > 10.0:
                                    _force_ok = False
                                    log(f'P{i}：回撤段且下一点为同位姿换姿——短直线让位 MoveJ 分支前视（v14w33c）。')
                            except Exception:
                                pass
                        if _force_ok:
                            lin_end_f, lin_detail_f = _linear_path_endpoint(q, target)
                            _lin_ok_f = (lin_end_f is not None
                                         and not _real_interfere_combo(lin_end_f)   # v14w26 组合禁区
                                         and (lookahead_ok is None or lookahead_ok(lin_end_f)))
                            if _lin_ok_f:
                                waypoints = _linear_waypoints(q, target)
                                if waypoints:
                                    end, method, fallback = lin_end_f, 'MoveL', True
                                    note = '短直线强制MoveL'
                                    forced_lin = True
                                    log(f'P{i}：短直线段（{_seg_mm_f:.1f}mm/姿态恒定）按工艺直走 MoveL（不尝试 MoveJ 弧）。')
                            elif lin_end_f is not None:
                                log(f'P{i}：短直线段直线末端无前视换向资格，回落 MoveJ 前视绑定。')
                            else:
                                log(f'P{i}：短直线段 MoveL 不可通行（{lin_detail_f}），回落 MoveJ 尝试。')
                        bound_applied = False
                        # v14j：前视绑定执行——本点是换向前夜：前视选出的构型若弧碰，不得退 MoveL
                        # （连续选解会静默锁回当前族，把死局推迟到换向步才爆——种子13 实证），
                        # 也不得由 v14c 救援收无前视资格的分支；只能换用其他前视合格分支直达，
                        # 全部失败则本构型判死、整段换种子重试。
                        if not forced_lin and lookahead_ok is not None and _movej_test_cached(q, end, 1) != 0:
                            detail_bound = _collision_details()
                            bound = None
                            for cand in sorted(_ik_branch_candidates(target, q),
                                               key=lambda c: sum((c[j]-q[j])**2 for j in range(6))):
                                if lookahead_ok(cand) and _movej_test_cached(q, cand, 1) == 0:
                                    bound = cand
                                    break
                            if bound is not None:
                                end, note, bound_applied = bound[:], '前视绑定避障直达', True
                                log(f'P{i}：前视构型弧碰（{detail_bound}），改用另一前视合格分支直达（前视绑定）。')
                            else:
                                raise ValueError(f'P{i}：MoveJ弧碰撞（{detail_bound}），其余前视合格分支均不可通行；'
                                                 '拒绝退 MoveL（连续选解会丢前视资格），本构型判死。')
                        # v14b：MoveJ 直达弧碰撞时，退回 v13 验证过的 MoveL 直线细分执行。
                        # v14w24：强制 MoveL 段不再尝试/回退 MoveJ（工艺直线优先）。
                        if not forced_lin and not bound_applied and _movej_test_cached(q, end, 1) != 0:
                            detail = _collision_details()
                            lin_end, lin_detail = _linear_path_endpoint(q, target)
                            if lin_end is None:
                                # v14c：直线也碰——枚举该目标全部 IK 分支找可通行 MoveJ（换构型救援）
                                # v14w33b：若下一点是【同位姿纯换姿】，优先选「下一点也能单条 MoveJ 贯通」
                                # 的救援分支（P6→P7 教训：P6 为自避碰选的分支对 P7 无路 ⇒ 49 跳细分拖死执行）。
                                _cands = sorted(_ik_branch_candidates(target, q),
                                                key=lambda c: sum((c[j] - q[j]) ** 2 for j in range(6)))
                                _nxt_pose = None
                                try:
                                    if i < len(records):
                                        _nr = records[i]
                                        if _nr['type'] == 'TCP' and not _nr.get('singular', False):
                                            _va = [float(v) for v in rec['values'][:6]]
                                            _vb = [float(v) for v in _nr['values'][:6]]
                                            if (all(abs(_va[k] - _vb[k]) < 1e-9 for k in range(3))
                                                    and any(abs(_va[k] - _vb[k]) > 1e-9 for k in range(3, 6))):
                                                _nxt_pose = fanuc_values_to_pose(*_nr['values'][:6])
                                except Exception:
                                    _nxt_pose = None
                                rescued = None
                                if _nxt_pose is not None:
                                    for cand in _cands:
                                        if _movej_test_cached(q, cand, 1) != 0:
                                            continue
                                        _ok_nxt = False
                                        for nb in _ik_branch_candidates(_nxt_pose, cand):
                                            if (_real_limit_ok(nb, lower, upper)
                                                    and not _real_interfere_combo(nb)
                                                    and _movej_test_cached(cand, nb, 1) == 0):
                                                _ok_nxt = True
                                                break
                                        if _ok_nxt:
                                            rescued = cand
                                            log(f'P{i}：下一点为同位姿换姿——救援分支带前视，选可与下一点单条 MoveJ 贯通的分支。')
                                            break
                                if rescued is None:
                                    for cand in _cands:
                                        if _movej_test_cached(q, cand, 1) == 0:
                                            rescued = cand
                                            break
                                if rescued is None:
                                    raise ValueError(f'P{i}：MoveJ弧碰撞（{detail}），且MoveL直线也失败：{lin_detail}；'
                                                     '该目标全部IK分支均不可通行。')
                                end, note = rescued[:], 'IK分支救援直达'
                                log(f'P{i}：最近解与直线均碰，切换IK分支救援成功。')
                            else:
                                # v14w33：同位姿/近零长（≤1mm）纯换姿段——MoveL 细分会把 90° 姿态差
                                # 切成数十跳小 MoveJ（10-21 P6→P7 实录 49 跳×每跳断连周期≈3s，
                                # 拖死执行）。优先搜无碰 MoveJ 分支单条直达（分支连续性绑死时
                                # 最近解弧碰≠无解）；搜不到再落回 MoveL 细分兜底。
                                # v14w34：_seg_mm_ro 必须是真实位置差——相对位姿平移模长在原地换姿
                                # 时被旋转杠杆放大（p−R·p，(0,-650,380) 处 90° 即 1064.8mm），
                                # 旧算式使 ≤1mm 门槛从未成立、两个搜索入口从未触发。
                                _pa = _trajectory_pose(q).Pos()
                                _pb = target.Pos()
                                _seg_mm_ro = math.sqrt(sum((_pa[_k] - _pb[_k]) ** 2 for _k in range(3)))
                                reorient_direct = None
                                if _seg_mm_ro <= 1.0:
                                    for cand in sorted(_ik_branch_candidates(target, q),
                                                       key=lambda c: sum((c[j]-q[j])**2 for j in range(6))):
                                        if (not _real_interfere_combo(cand)
                                                and _real_limit_ok(cand, lower, upper)
                                                and (lookahead_ok is None or lookahead_ok(cand))
                                                and _movej_test_cached(q, cand, 1) == 0):
                                            reorient_direct = cand
                                            break
                                if reorient_direct is not None:
                                    end, note = reorient_direct[:], '同位姿换姿MoveJ直达'
                                    method, fallback = 'MoveJ', False
                                    waypoints = []
                                    log(f'P{i}：同位姿换姿——MoveL 细分会碎成数十小段，改用无碰 MoveJ 分支单条直达。')
                                elif _seg_mm_ro <= 1.0 and plan and rec['type'] == 'TCP' and i >= 2:
                                    # v14w33d：回改上一步（已入计划、未执行）为可与本点单条 MoveJ 贯通的
                                    # 分支——上一步若走最近解直达/救援，其分支未必对本点有路（P6→P7 实录）。
                                    # 改关节目标后两跳路径均当场重检，证书完整。
                                    _prev_step = plan[-1]
                                    _prev_q = _prev_step['joints']
                                    _prev_prev = plan[-2]['joints'] if len(plan) >= 2 else saved
                                    _prev_pose = fanuc_values_to_pose(*records[i - 2]['values'][:6])
                                    reorient_direct = None
                                    for c6 in sorted(_ik_branch_candidates(_prev_pose, _prev_prev),
                                                     key=lambda c: sum((c[k] - _prev_q[k]) ** 2 for k in range(6))):
                                        if _real_interfere_combo(c6) or not _real_limit_ok(c6, lower, upper):
                                            continue
                                        if _movej_test_cached(_prev_prev, c6, 1) != 0:
                                            continue
                                        for c7 in sorted(_ik_branch_candidates(target, c6),
                                                         key=lambda c: sum((c[k] - c6[k]) ** 2 for k in range(6))):
                                            if _real_interfere_combo(c7) or not _real_limit_ok(c7, lower, upper):
                                                continue
                                            if lookahead_ok is not None and not lookahead_ok(c7):
                                                continue
                                            if _movej_test_cached(c6, c7, 1) != 0:
                                                continue
                                            _prev_step['joints'] = c6[:]
                                            reorient_direct = c7
                                            break
                                        if reorient_direct is not None:
                                            break
                                    if reorient_direct is not None:
                                        end, note = reorient_direct[:], '同位姿换姿MoveJ直达'
                                        method, fallback = 'MoveJ', False
                                        waypoints = []
                                        log(f'P{i}：回改上一步分支后，本点取得单条 MoveJ 直达（两跳均重检无碰）。')
                                if reorient_direct is not None:
                                    pass   # 已在上方处理
                                else:
                                    waypoints = _linear_waypoints(q, target)
                                    if not waypoints:
                                        raise ValueError(f'P{i}：MoveJ弧碰撞（{detail}），MoveL细分采样失败，拒绝。')
                                    end, method, fallback = lin_end, 'MoveL', True
                                    note = 'MoveJ弧碰退回MoveL细分'
                                    log(f'P{i}：MoveJ弧碰撞（{detail}），改走 MoveL 直线细分（{len(waypoints)} 途经点）。')
                    if not all(lower[j] <= end[j] <= upper[j] for j in range(6)):
                        raise ValueError(f'P{i}：关节超限，J6目标={end[5]:.3f}°。')
                    if method == 'MoveJ' and _movej_test_cached(q, end, 1) != 0:
                        # v14e：普通TCP点最后一级救援——v13 遗产 _obstacle_joint_target
                        # （21候选、肘高排序、限TCP偏离）选避障构型，TCP仿真靠它在同一站过关。
                        try:
                            end = _obstacle_joint_target(q, rec['values'], max_deviation, log)
                            note = '避障选解直达'
                        except ValueError:
                            raise ValueError(f'P{i}：MoveJ路径检查失败（含避障选解）：' + _collision_details())
                        if _movej_test_cached(q, end, 1) != 0:
                            raise ValueError(f'P{i}：MoveJ路径检查失败：' + _collision_details())
                    # v15.22: try the equivalent J6 winding before committing a long fallback.
                    if not rec.get('singular') and 170.0 <= end[5] <= 360.0 and i < len(records) and any(r.get('singular') and not r.get('spin360') for r in records[max(0,i-2):min(len(records),i+2)]):
                        adjusted = end[:]
                        adjusted[5] -= 360.0
                        if (_real_limit_ok(adjusted, lower, upper) and not _real_interfere_combo(adjusted)
                                and _movej_test_cached(q, adjusted, 1) == 0):
                            if method == 'MoveJ' or (waypoints and norm((target * invH(_trajectory_pose(q))).Pos()) > MOVL_DIRECT_MAX_MM):
                                log(f'P{i}：J6同角分支 {end[5]:.3f}→{adjusted[5]:.3f}°，MoveJ路径已复核。')
                                end, method, waypoints = adjusted, 'MoveJ', []
                    # v14w25：J6 恰=±360 边界值被控制器 -40006 拒收（10-15 17:26/17:33 实录）。
                    # v14w32：±359.999 内推仍防不住「J6 单轴被丢弃」（10-21 P4 实证：J1~J5 全到、
                    # J6 纹丝停在 180、误差 180°）——改为换 (−180,180] 同角表示（359.999→−0.001），
                    # J6 彻底离开 ±360 邻域。换表示会翻转 MoveJ 弧方向 ⇒ 必须重检路径，不过即报规划错误。
                    # spin360/多圈值（|J6|>360.001）不在此列，防绞坏自转语义。
                    if 359.0 <= abs(end[5]) <= 360.001 and not rec.get('spin360'):
                        _j6n = end[5] - math.copysign(360.0, end[5])
                        log(f'P{i}：J6={end[5]:.3f}° 进入 ±360 一度防护区，换同角表示 {_j6n:.3f}°（v15.22：359.45实测未执行，换向后重检路径）。')
                        if waypoints:
                            raise ValueError(f'P{i}：J6进入±360的一度防护区，连续直线需换分支重新认证。')
                        end[5] = _j6n
                        if rec.get('singular'):
                            delta = int(round(end[5] - q[5]))
                        for _wp in waypoints:
                            if abs(_wp[5]) >= 359.999 and abs(_wp[5]) <= 360.001:
                                _wp[5] = _wp[5] - math.copysign(360.0, _wp[5])
                        if method == 'MoveJ' and _movej_test_cached(q, end, 1) != 0:
                            raise ValueError(f'P{i}：J6 换同角表示后 MoveJ 路径碰撞：' + _collision_details())
                    # v14w26：解落入实机自干涉组合区（J4×J5，-40006）——MoveJ 解自动换无碰安全
                    # 分支直达；直线段落区（强制/兜底）整段换种子；无安全分支则判死。
                    if _real_interfere_combo(end):
                        if method == 'MoveJ' and rec['type'] == 'TCP' and not rec.get('singular', False):
                            rescued_if = None
                            for cand_if in sorted(_ik_branch_candidates(target, q),
                                                   key=lambda c: sum((c[j]-q[j])**2 for j in range(6))):
                                if (_real_limit_ok(cand_if, lower, upper)
                                        and not _real_interfere_combo(cand_if)
                                        and _movej_test_cached(q, cand_if, 1) == 0):
                                    rescued_if = cand_if
                                    break
                            if rescued_if is None:
                                raise ValueError(f'P{i}：全部无碰分支均落入实机自干涉组合区'
                                                 f'（|J4|>{REAL_INTERFERE_J4_MAX:.0f} 且 |J5|>{REAL_INTERFERE_J5_MIN:.0f}，-40006 实录区），本构型判死。')
                            log(f'P{i}：预选解落入实机自干涉组合区（J4={end[3]:.1f}°, J5={end[4]:.1f}°），换安全分支直达。')
                            end = rescued_if[:]
                            note = '自干涉安全分支直达'
                        else:
                            raise ValueError(f'P{i}：该步解落入实机自干涉组合区（J4={end[3]:.1f}°, J5={end[4]:.1f}°），换种子重试。')
                    plan.append(dict(method=method, joints=end[:], special=rec.get('singular', False), fallback=False,
                                     rewinds=rewinds, j6_delta=delta,
                                     waypoints=waypoints, p2p_note=note))
                    q = end[:]
                if _continuous_profile_active:
                    previous = saved
                    for number, step in enumerate(plan, 1):
                        if step.get('waypoints'):
                            rel = _trajectory_pose(step['joints']) * invH(_trajectory_pose(previous))
                            if (step['method'] != 'MoveL' or norm(rel.Pos()) > MOVL_DIRECT_MAX_MM
                                    or pose_angle(rel) > math.radians(.5)):
                                raise ValueError(f'P{number}将退回{len(step["waypoints"])}段停走，换入口分支重试。')
                        previous = step['joints']
                log('逐段规划完成，开始整段碰撞复核（1mm/1°采样，请稍候）…')
                _verify_obstacle_plan(saved, plan)
                _certify_continuous_direct(records, saved, plan, log)
                _preferred_seed = (seed_context, seed)
                log(f'P2P+奇异点整段路径预检通过：{len(plan)}点。')
                return plan
            except ValueError as exc:
                last_seed_error = exc
                log(f'种子 {seed_rank}/{len(seeds)} 在此构型失败（{exc}），换下一构型整段重试…')
        if last_seed_error is not None:
            raise last_seed_error
    finally:
        _continuous_profile_active = False
        robot.setJoints(saved)
        RDK.Render(True)

root = tk.Tk()
root.title("RoboDK - 机械臂运动控制（P2P v15.22）")
root.geometry("1200x750")
root.resizable(True, True)

tk.Label(root, text="Dobot CR5 运动控制", font=("Microsoft YaHei", 16, "bold")).pack(pady=10)

notebook = ttk.Notebook(root)
notebook.pack(fill=tk.BOTH, expand=True, padx=10, pady=5)

# ---- 选项卡 1：单点运动 ----
tab_single = ttk.Frame(notebook)
notebook.add(tab_single, text="单点运动")

frame_coord = tk.LabelFrame(tab_single, text="目标 TCP（Fanuc 格式）")
frame_coord.pack(fill=tk.X, padx=10, pady=10)

names = ["X (mm)", "Y (mm)", "Z (mm)", "Rx (deg)", "Ry (deg)", "Rz (deg)"]
defaults = ["0.000", "-241.500", "1047.000", "-90.000", "0.000", "180.000"]
entries_single = []

for i in range(6):
    tk.Label(frame_coord, text=names[i]).grid(row=0, column=i*2, padx=5, pady=10)
    e = tk.Entry(frame_coord, width=12)
    e.insert(0, defaults[i])
    e.grid(row=0, column=i*2+1, padx=5, pady=10)
    entries_single.append(e)

frame_mtype = tk.Frame(tab_single)
frame_mtype.pack(fill=tk.X, padx=10, pady=5)
move_type = tk.StringVar(value="MoveL")
tk.Radiobutton(frame_mtype, text="MoveL (直线)", variable=move_type, value="MoveL").pack(side=tk.LEFT, padx=10)
tk.Radiobutton(frame_mtype, text="MoveJ (关节)", variable=move_type, value="MoveJ").pack(side=tk.LEFT, padx=10)

btn_single_frame = tk.Frame(tab_single)
btn_single_frame.pack(fill=tk.X, padx=10, pady=5)

def _read_current():
    read_current(entries_single)
def _fill_current():
    fill_current(entries_single)
def _check_ik():
    check_ik_single(entries_single)
def _exec_single():
    execute_single(entries_single, move_type.get())

tk.Button(btn_single_frame, text="读取当前 TCP", command=_read_current, width=15).pack(side=tk.LEFT, padx=3)
tk.Button(btn_single_frame, text="当前 TCP -> 输入框", command=_fill_current, width=20).pack(side=tk.LEFT, padx=3)
tk.Button(btn_single_frame, text="检测可达性", command=_check_ik, width=15, bg="#2196F3", fg="white").pack(side=tk.LEFT, padx=3)
tk.Button(btn_single_frame, text="执行运动", command=_exec_single, width=20,
          font=("Microsoft YaHei", 10, "bold"), bg="#4CAF50", fg="white").pack(side=tk.LEFT, padx=3)


# ---- 选项卡 2：目标关节运动（实机） ----
tab_joint = ttk.Frame(notebook)
notebook.add(tab_joint, text="目标关节运动")

frame_joint = tk.LabelFrame(tab_joint, text="目标关节（deg）")
frame_joint.pack(fill=tk.X, padx=10, pady=10)

joint_names = ["J1 (deg)", "J2 (deg)", "J3 (deg)", "J4 (deg)", "J5 (deg)", "J6 (deg)"]
joint_defaults = ["0.000", "0.000", "0.000", "0.000", "0.000", "0.000"]
entries_joint = []

for i in range(6):
    tk.Label(frame_joint, text=joint_names[i]).grid(row=0, column=i*2, padx=5, pady=10)
    e = tk.Entry(frame_joint, width=12)
    e.insert(0, joint_defaults[i])
    e.grid(row=0, column=i*2+1, padx=5, pady=10)
    entries_joint.append(e)

btn_joint_frame = tk.Frame(tab_joint)
btn_joint_frame.pack(fill=tk.X, padx=10, pady=8)

def _read_current_joint_values():
    read_current_joints(entries_joint)

def _fill_current_joints():
    fill_current_joints(entries_joint)

def _exec_joint():
    execute_joint_target(entries_joint)

def _zero_joints():
    clear_joint_target(entries_joint)

tk.Button(btn_joint_frame, text="读取当前关节", command=_read_current_joint_values, width=14).pack(side=tk.LEFT, padx=3)
tk.Button(btn_joint_frame, text="当前关节 -> 输入框", command=_fill_current_joints, width=20).pack(side=tk.LEFT, padx=3)
tk.Button(btn_joint_frame, text="执行指定关节 MoveJ", command=_exec_joint, width=24,
          font=("Microsoft YaHei", 10, "bold"), bg="#FF9800", fg="white").pack(side=tk.LEFT, padx=3)
tk.Button(btn_joint_frame, text="清零", command=_zero_joints, width=10).pack(side=tk.LEFT, padx=3)

tk.Label(tab_joint,
         text="输入 J1~J6 目标角度（deg）；完整关节路径预检通过后才发送实机 MoveJ。",
         fg="#555555").pack(anchor=tk.W, padx=15, pady=5)
tk.Label(tab_joint,
         text="安全提示：首次测试建议只改变一个关节、改变 5~10°，确认方向和角度定义正确后再进行大角度运动。",
         fg="#C62828").pack(anchor=tk.W, padx=15, pady=2)

# ---- 选项卡 3：连续运动 ----
tab_traj = ttk.Frame(notebook)
notebook.add(tab_traj, text="连续运动")

frame_traj_input = tk.LabelFrame(
    tab_traj,
    text="连续运动点输入：每次输入 1 个 TCP 点或 1 组关节角度，点击“检查并加入”"
)
frame_traj_input.pack(fill=tk.X, padx=10, pady=10)

type_frame = tk.Frame(frame_traj_input)
type_frame.pack(fill=tk.X, padx=8, pady=5)

tk.Label(type_frame, text="点类型：").pack(side=tk.LEFT, padx=3)

traj_type = tk.StringVar(value="TCP")
tk.Radiobutton(
    type_frame, text="TCP（X,Y,Z,Rx,Ry,Rz）",
    variable=traj_type, value="TCP"
).pack(side=tk.LEFT, padx=8)

tk.Radiobutton(
    type_frame, text="关节（J1~J6）",
    variable=traj_type, value="JOINT"
).pack(side=tk.LEFT, padx=8)

traj_names_tcp = ["X", "Y", "Z", "Rx", "Ry", "Rz"]
traj_names_joint = ["J1", "J2", "J3", "J4", "J5", "J6"]

traj_entries = []

# ---- 末端特异点设置 ----
singular_var = tk.BooleanVar(value=False)
j6_direction_var = tk.IntVar(value=180)

singular_frame = tk.Frame(frame_traj_input)
singular_frame.pack(fill=tk.X, padx=8, pady=3)

tk.Checkbutton(
    singular_frame,
    text="末端特异点（跳过IK，仅J6转动）",
    variable=singular_var
).pack(side=tk.LEFT, padx=3)

tk.Label(singular_frame, text="J6方向：").pack(side=tk.LEFT, padx=(15, 3))
tk.Radiobutton(singular_frame, text="+180°", variable=j6_direction_var, value=180).pack(side=tk.LEFT, padx=3)
tk.Radiobutton(singular_frame, text="-180°", variable=j6_direction_var, value=-180).pack(side=tk.LEFT, padx=3)
spin_var = tk.BooleanVar(value=False)
tk.Checkbutton(singular_frame, text="J6自转360°（第二类，六维与前点相同）", variable=spin_var).pack(side=tk.LEFT, padx=3)

# 输入框单独放在 grid 子容器中。
# frame_traj_input 本身使用 pack 管理子控件，不能再直接对它的子控件使用 grid。
traj_value_frame = tk.Frame(frame_traj_input)
traj_value_frame.pack(fill=tk.X, padx=8, pady=5)

for i in range(6):
    tk.Label(
        traj_value_frame,
        text=traj_names_tcp[i]
    ).grid(row=0, column=i * 2, padx=3, pady=8)

    e = tk.Entry(traj_value_frame, width=12)
    e.grid(row=0, column=i * 2 + 1, padx=4, pady=8)
    traj_entries.append(e)

# 默认先按 TCP 输入显示
tcp_defaults = ["0.000", "-241.500", "1047.000", "-90.000", "0.000", "180.000"]
for e, val in zip(traj_entries, tcp_defaults):
    e.insert(0, val)


def _update_traj_labels_and_defaults():
    """切换 TCP/关节输入时，更新标签和默认值。"""
    names = traj_names_tcp if traj_type.get() == "TCP" else traj_names_joint
    defaults = (
        tcp_defaults
        if traj_type.get() == "TCP"
        else ["0.000"] * 6
    )

    for i, e in enumerate(traj_entries):
        # grid 上的 Label 位于当前列
        for widget in traj_value_frame.grid_slaves(row=0, column=i * 2):
            widget.configure(text=names[i])

        e.delete(0, tk.END)
        e.insert(0, defaults[i])


tk.Radiobutton(
    type_frame, text="TCP（X,Y,Z,Rx,Ry,Rz）",
    variable=traj_type, value="TCP",
    command=_update_traj_labels_and_defaults
).pack_forget()

# 重新建立带 command 的两个单选按钮
for widget in list(type_frame.pack_slaves()):
    if isinstance(widget, tk.Radiobutton):
        widget.destroy()

tk.Radiobutton(
    type_frame, text="TCP（X,Y,Z,Rx,Ry,Rz）",
    variable=traj_type, value="TCP",
    command=_update_traj_labels_and_defaults
).pack(side=tk.LEFT, padx=8)

tk.Radiobutton(
    type_frame, text="关节（J1~J6）",
    variable=traj_type, value="JOINT",
    command=_update_traj_labels_and_defaults
).pack(side=tk.LEFT, padx=8)

btn_traj_input = tk.Frame(tab_traj)
btn_traj_input.pack(fill=tk.X, padx=10, pady=3)

tk.Button(
    btn_traj_input,
    text="检查并加入当前点",
    command=add_and_check_trajectory_point,
    width=22,
    bg="#2196F3",
    fg="white",
    font=("Microsoft YaHei", 10, "bold")
).pack(side=tk.LEFT, padx=3)

tk.Button(
    btn_traj_input,
    text="读取当前TCP并写入",
    command=read_current_tcp_to_traj,
    width=20
).pack(side=tk.LEFT, padx=3)

tk.Button(
    btn_traj_input,
    text="读取当前关节并写入",
    command=read_current_joints_to_traj,
    width=20
).pack(side=tk.LEFT, padx=3)

tk.Button(
    btn_traj_input,
    text="清空当前输入",
    command=clear_trajectory_input,
    width=16
).pack(side=tk.LEFT, padx=3)

tk.Label(
    tab_traj,
    text="加入点时检查格式并保留关节圈数；执行前再进行整段限位、台子和地面碰撞检查。",
    fg="#555555"
).pack(anchor=tk.W, padx=15, pady=3)

frame_record = tk.LabelFrame(
    tab_traj,
    text="已检查通过的连续运动点（按加入顺序执行，可混合 TCP / 关节点）"
)
frame_record.pack(fill=tk.BOTH, expand=True, padx=10, pady=8)

record_text = tk.Text(frame_record, font=("Consolas", 10), height=10)
record_text.pack(fill=tk.BOTH, expand=True, padx=5, pady=5)

btn_record_frame = tk.Frame(tab_traj)
btn_record_frame.pack(fill=tk.X, padx=10, pady=4)

tk.Button(
    btn_record_frame, text="删除最后一点",
    command=delete_last_record, width=15
).pack(side=tk.LEFT, padx=3)

tk.Button(
    btn_record_frame, text="清空全部点",
    command=clear_records, width=15
).pack(side=tk.LEFT, padx=3)

tk.Button(
    btn_record_frame, text="导入轨迹",
    command=import_trajectory, width=14
).pack(side=tk.LEFT, padx=3)

tk.Button(
    btn_record_frame, text="执行整段连续运动",
    command=execute_recorded_trajectory,
    width=24,
    font=("Microsoft YaHei", 10, "bold"),
    bg="#4CAF50", fg="white"
).pack(side=tk.LEFT, padx=3)

tk.Label(
    tab_traj,
    text="执行前按实机当前关节完成台子/地面预检；仅执行已验证方案。驱动报断连时复核实际到位；未到位或其他异常时中止。",
    fg="#555555"
).pack(anchor=tk.W, padx=15, pady=4)

real_deviation_var = tk.StringVar(value="500.0")
frame_deviation = tk.Frame(root)
frame_deviation.pack(fill=tk.X, padx=10, pady=3)
tk.Label(frame_deviation, text="预检MoveJ兜底最大TCP偏离(mm)：").pack(side=tk.LEFT)
tk.Entry(frame_deviation, textvariable=real_deviation_var, width=10).pack(side=tk.LEFT)
tk.Label(frame_deviation, text="默认500：与TCP仿真/轨迹7~11验证口径一致；实机速度10 mm/s（v14w25 调慢）").pack(side=tk.LEFT, padx=8)

# v14w24：法兰补偿MOVL 默认开启，勾选框移除（工艺定型）。v14l 实机判决驱动 MOVL 无工具
# 补偿（按法兰执行，无补偿直发已拉黑勿回归）；v14p 将错就错把法兰位姿当笛卡尔目标直发，
# 法兰被精确送达→物理尖端走在认证直线上。v14w36/37：位姿由调用方自算 invH(PoseFrame)*SolveFK
# （动画=认证直线，根治关节弧假碰撞冻死），发送窗口配单位变换（校验/数字=法兰空间）。
# 适用：MoveL 细分段≤210mm 且姿态恒定（v14w35 门禁）；规划/预检/几何零改动；失败指纹照旧即停；净化失败自动回落细分。
real_movldirect_var = tk.BooleanVar(value=True)   # 仅保留变量接口（执行入口读取）；无 GUI 控件

# ---- 日志区 ----
frame_log = tk.LabelFrame(root, text="日志")
frame_log.pack(fill=tk.BOTH, expand=True, padx=10, pady=5)

text_log = scrolledtext.ScrolledText(frame_log, font=("Consolas", 10), height=8)
text_log.pack(fill=tk.BOTH, expand=True, padx=5, pady=5)

# ============================================================
# 启动
# ============================================================
log("机器人: " + robot.Name())
log("程序就绪。" + LOG_VERSION + " ｜ 模式：RUNMODE_RUN_ROBOT + robot.Connect() ｜ 文件日志：" + LOG_PATH)
_ensure_canonical_tool()   # v14w17：启动守护（覆盖"加载了带归零工具的存档"场景）
log("单点：输入坐标 -> 检测可达性 -> 执行 MoveL/MoveJ")
log("目标关节：输入 J1~J6 -> 实机 MoveJ（不经过 TCP/Fanuc 转换和 IK）")
log("连续运动（P2P v15.22）：修改点位后仍启用分支搜索、防停走及逐段重新认证；无法认证的直线在发送运动前停止；130mm TCP。")

def _log_pump():
    try:
        while True:
            text_log.insert(tk.END, _log_queue.get_nowait() + NL)
            text_log.see(tk.END)
    except Exception:
        pass
    root.after(100, _log_pump)


_close_requested = False


def _idle_tool_guard():
    if not _real_running and not _tool_window_depth:
        try:
            if _same_tool_pose(robot.PoseTool(), eye(4)):
                _ensure_canonical_tool()
            if _close_requested:
                root.destroy()
                return
        except Exception as exc:
            _file_log('工具空闲守护失败：' + str(exc))
    root.after(1000, _idle_tool_guard)


def _on_close():
    global _close_requested
    if _real_running:
        _close_requested = True
        log('已请求关闭：等待当前任务结束并恢复 TCP 后关闭窗口，继续保留到位监控。')
        return
    _ensure_canonical_tool()
    root.destroy()


root.protocol('WM_DELETE_WINDOW', _on_close)
root.after(100, _log_pump)
root.after(1000, _idle_tool_guard)
_start_heartbeat()
try:
    root.mainloop()
except BaseException:
    import traceback
    _file_log('FATAL mainloop: ' + traceback.format_exc())
    raise

--- program 轨迹17_仿真27点 (robot Dobot CR5) ---
  设置参考: Dobot CR5 Base_控制器对齐
  设置工具 at (0, 0, 130) mm
  MoveJ (回放17_27点_00) to (0.81, -375.18, 1048.46) mm, rotated rx -89.77 ry 0 rz 179.86 deg; joints [0, 0, 0, 0, 0, 0]
  MoveJ (回放17_27点_01) to (500, 0, 460) mm, rotated rx 180 ry 0 rz 0 deg; joints [15.907, -63.543, 66.599, -93.225, 90.382, -73.897]
  MoveJ (回放17_27点_02) to (0, -551.1, 420) mm, rotated rx -90 ry 0 rz -180 deg; joints [64.021, 6.446, 132.247, -138.394, -63.355, -0.324]
  MoveL (回放17_27点_03) to (120, -551.1, 420) mm, rotated rx -90 ry 0 rz -180 deg; joints [86.577, 9.276, 128.708, -137.798, -85.916, -0.207]
  MoveJ (回放17_27点_04) to (120, -551.1, 420) mm, rotated rx 90 ry 0 rz 0 deg; joints [86.577, 9.276, 128.708, -137.798, -85.916, 179.793]
  MoveL (回放17_27点_05) to (20, -551.13, 420) mm, rotated rx 90 ry 0 rz 0 deg; joints [67.69, 6.533, 132.142, -138.399, -67.023, 179.697]
  MoveL (回放17_27点_06) to (-135, -551.17, 420) mm, rotated rx 90 ry 0 rz 0 deg; joints [43.2, 9.991, 127.778, -137.308, -42.54, 179.533]
  MoveJ (回放17_27点_07) to (0, -516.17, 420) mm, rotated rx 90 ry 0 rz 0 deg; joints [60.482, 1.539, 137.799, -138.995, -59.811, 179.613]
  MoveJ (回放17_27点_08) to (0, -516.17, 420) mm, rotated rx 180 ry 0 rz 0 deg; joints [-73.904, -4.388, -72.292, -13.492, 89.709, 195.818]
  MoveL (回放17_27点_09) to (0, -538.81, 420) mm, rotated rx -180 ry 0 rz 0 deg; joints [-74.605, -7.638, -68.632, -13.901, 89.734, 195.121]
  MoveL (回放17_27点_10) to (-125, -538.82, 420) mm, rotated rx -180 ry 0 rz 0 deg; joints [-88.08, -9.727, -66.162, -14.284, 89.751, 181.651]
  MoveJ (回放17_27点_11) to (-125, -538.82, 420) mm, rotated rx -180 ry 0 rz 180 deg; joints [-88.08, -9.727, -66.162, -14.284, 89.751, 1.651]
  MoveL (回放17_27点_12) to (0, -538.81, 420) mm, rotated rx 180 ry 0 rz -180 deg; joints [-74.605, -7.638, -68.632, -13.901, 89.734, 15.121]
  MoveL (回放17_27点_13) to (125, -538.81, 420) mm, rotated rx 180 ry 0 rz -180 deg; joints [-61.957, -9.725, -66.163, -14.283, 89.751, 27.774]
  MoveJ (回放17_27点_14) to (40, -503.8, 420) mm, rotated rx 90 ry 0 rz 90 deg; joints [54.027, 22.646, 68.332, 89.289, -36.384, -0.204]
  MoveL (回放17_27点_15) to (30, -538.8, 420) mm, rotated rx 90 ry 0 rz 90 deg; joints [55.298, 28.251, 59.827, 92.253, -35.079, -0.283]
  MoveJ (回放17_27点_16) to (40, -503.81, 420) mm, rotated rx 131.17 ry 90 rz 131.17 deg; joints [54.027, 22.647, 68.33, 89.29, -36.384, -90.204]
  MoveL (回放17_27点_17) to (30, -538.81, 420) mm, rotated rx 0 ry 90 rz 0 deg; joints [55.299, 28.252, 59.825, 92.253, -35.078, -90.283]
  MoveJ (回放17_27点_18) to (40, -503.81, 420) mm, rotated rx -131.17 ry -90 rz -48.83 deg; joints [54.028, 22.648, 68.329, 89.29, -36.383, -270.205]
  MoveL (回放17_27点_19) to (30, -538.81, 420) mm, rotated rx 0 ry -90 rz -180 deg; joints [55.299, 28.253, 59.824, 92.254, -35.078, -270.283]
  MoveJ (回放17_27点_20) to (50, -503.8, 420) mm, rotated rx -88.93 ry -59.66 rz -90.94 deg; joints [54.921, 22.39, 69.063, 89.747, -35.48, -240.633]
  MoveL (回放17_27点_21) to (40, -538.8, 420) mm, rotated rx -88.93 ry -59.66 rz -90.94 deg; joints [56.146, 27.979, 60.611, 92.705, -34.223, -240.749]
  MoveL (回放17_27点_22) to (40, -498.8, 420) mm, rotated rx -88.93 ry -59.66 rz -90.94 deg; joints [53.698, 22.211, 69.324, 89.629, -36.704, -240.588]
  MoveJ (回放17_27点_23) to (50, -503.8, 420) mm, rotated rx 90 ry 0 rz 90 deg; joints [54.925, 22.121, 69.098, 89.049, -35.489, -0.205]
  MoveJ (回放17_27点_24) to (40, -504.28, 420) mm, rotated rx -88.93 ry 59.66 rz -90.94 deg; joints [53.576, 21.931, 69.73, 89.548, -34.985, -121.311]
  MoveL (回放17_27点_25) to (40, -539.28, 420) mm, rotated rx -88.93 ry 59.66 rz -90.94 deg; joints [55.751, 26.938, 62.23, 92.167, -32.782, -121.461]
  MoveL (回放17_27点_26) to (40, -499.28, 420) mm, rotated rx -88.93 ry 59.66 rz -90.94 deg; joints [53.243, 21.24, 70.728, 89.225, -35.321, -121.29]
  MoveJ (回放17_27点_27) to (-600, 0, 460) mm, rotated rx 180 ry 0 rz -90 deg; joints [-13.36, 19.281, 46.973, 23.918, -90.105, -193.743]

--- Python program CR5_零位到P1_上传 ---
"""RoboDK station macro that uploads the reviewed P1 project on button click."""
import errno
import hashlib
from pathlib import Path
import re
import socket
import sys
import threading
import tkinter as tk
from tkinter import ttk
import uuid

WORKSPACE = Path(r"D:\mydata\glm-workplace")
PROJECT_NAME = "CR5_Traj17_ZeroToP1"
PROJECT = WORKSPACE / "sim_scripts/rdk_station_dump/cr5_controller_deployment_check" / PROJECT_NAME
REMOTE_ROOT = "/dobot/userdata/project/project"
FILES = ("prj.json", "global.lua", "point.json", "point.json.lua", "src0.lua")
EXPECTED = {'global.lua': '01ba4719c80b6fe911b091a7c05124b64eeece964e09c058ef8f9805daca546b', 'point.json': '37517e5f3dc66819f61f5a7bb8ace1921282415f10551d2defa5c3eb0985b570', 'point.json.lua': 'e3b0c44298fc1c149afbf4c8996fb92427ae41e4649b934ca495991b7852b855', 'prj.json': '14f1471434bc39ae6f11944fdff35eff23d14d9e65682650c694a0375f86ce9c', 'src0.lua': 'c66c50b254430aadf534d1c7742c74fdf04aac4593f4b490c3d254d51c0740ae'}


def exists(sftp, path):
    try:
        sftp.stat(path)
    except OSError as error:
        if error.errno == errno.ENOENT:
            return False
        raise
    return True


def upload(allow_create=True):
    sys.path.insert(0, str(WORKSPACE / "tools"))
    import rssh
    import paramiko

    content = {name: (PROJECT / name).read_bytes() for name in FILES}
    if {name: hashlib.sha256(data).hexdigest() for name, data in content.items()} != EXPECTED:
        raise RuntimeError("本地工程与已核对版本不一致。")
    target = REMOTE_ROOT + "/" + PROJECT_NAME
    pending = REMOTE_ROOT + "/." + PROJECT_NAME + "_" + uuid.uuid4().hex
    client = paramiko.SSHClient()
    client.set_missing_host_key_policy(paramiko.AutoAddPolicy())
    try:
        client.connect(rssh.HOST, username=rssh.USER, password=rssh.PASS,
                       timeout=8, allow_agent=False, look_for_keys=False)
        with client.open_sftp() as sftp:
            sftp.get_channel().settimeout(8)

            def verify(folder):
                for name, data in content.items():
                    with sftp.open(folder + "/" + name, "rb") as file:
                        if file.read() != data:
                            raise RuntimeError("回读不一致：" + name)

            if exists(sftp, target):
                verify(target)
                return "工程已在控制器，文件回读一致。"
            if not allow_create:
                raise RuntimeError("请先上传工程。")
            sftp.mkdir(pending)
            try:
                for name, data in content.items():
                    with sftp.open(pending + "/" + name, "wb") as file:
                        file.write(data)
                verify(pending)
                sftp.rename(pending, target)
            except Exception:
                if exists(sftp, pending):
                    for name in FILES:
                        path = pending + "/" + name
                        if exists(sftp, path):
                            sftp.remove(path)
                    sftp.rmdir(pending)
                raise
            verify(target)
            return "上传完成，控制器端 5 个文件回读一致。"
    finally:
        client.close()


def start_project():
    upload(allow_create=False)
    import rssh

    def command(connection, request):
        connection.sendall(request.encode("ascii"))
        data = b""
        while b";" not in data:
            chunk = connection.recv(4096)
            if not chunk:
                raise RuntimeError("命令口无应答，请确认 RoboDK 驱动已断开。")
            data += chunk
        return data.decode("ascii", errors="replace")

    def values(reply):
        match = re.match(r"^\s*0,\{([^}]*)\}", reply)
        if not match:
            raise RuntimeError("控制器拒绝查询：" + reply)
        return [float(value) for value in match.group(1).split(",") if value]

    with socket.create_connection((rssh.HOST, 29999), timeout=4) as connection:
        if values(command(connection, "RobotMode()")) != [5.0]:
            raise RuntimeError("控制器未处于已使能待机状态。")
        axes = values(command(connection, "GetAngle()"))
        if len(axes) != 6 or not all(abs(angle) <= 0.05 for angle in axes):
            raise RuntimeError("六轴起始角度不在零位容差内。")
        connection.sendall(("RunScript(" + PROJECT_NAME + ")").encode("ascii"))
        try:
            reply = connection.recv(4096).decode("ascii", errors="replace")
        except OSError:
            return "启动命令已发送，应答未确认。请查看控制器状态，避免重复点击。"
        if not reply:
            return "启动命令已发送，应答未确认。请查看控制器状态，避免重复点击。"
        if not re.match(r"^\s*0,", reply):
            raise RuntimeError("控制器拒绝启动：" + reply)
    return "控制器已接受启动命令。请观察零位→P1 的运动和到位状态。"


def run_action(action, pending, lock_start=False):
    button.configure(state="disabled")
    start_button.configure(state="disabled")
    status.set(pending)

    def worker():
        try:
            message = action()
            locked = lock_start
        except Exception as error:
            message = "操作未完成：" + str(error)
            locked = False
        try:
            window.after(0, finish, message, locked)
        except (RuntimeError, tk.TclError):
            pass

    threading.Thread(target=worker, daemon=False).start()


def finish(message, locked):
    status.set(message)
    button.configure(state="normal")
    if not locked:
        start_button.configure(state="normal")


if __name__ == "__main__":
    window = tk.Tk()
    window.title("CR5 零位→P1 工程上传")
    status = tk.StringVar(value="等待上传。上传与启动分开。点击启动会使实机从零位移动到 P1。")
    ttk.Label(window, text=PROJECT_NAME, padding=12).pack()
    button = ttk.Button(window, text="上传到控制器", command=lambda: run_action(upload, "正在上传并校验…"))
    button.pack(pady=5)
    start_button = ttk.Button(window, text="启动零位→P1（实机运动）",
                              command=lambda: run_action(start_project, "核对工程及控制器状态…", True))
    start_button.pack(pady=5)
    ttk.Label(window, textvariable=status, wraplength=480, padding=12).pack()
    window.mainloop()

--- Python program CR5_首段MoveL_上传 ---
"""RoboDK station macro that uploads the reviewed P1 project on button click."""
import errno
import hashlib
from pathlib import Path
import re
import socket
import sys
import threading
import tkinter as tk
from tkinter import ttk
import uuid

WORKSPACE = Path(r"D:\mydata\glm-workplace")
PROJECT_NAME = "CR5_Traj17_ZeroToFirstMoveL"
PROJECT = WORKSPACE / "sim_scripts/rdk_station_dump/cr5_controller_deployment_check" / PROJECT_NAME
REMOTE_ROOT = "/dobot/userdata/project/project"
FILES = ("prj.json", "global.lua", "point.json", "point.json.lua", "src0.lua")
EXPECTED = {'global.lua': '01ba4719c80b6fe911b091a7c05124b64eeece964e09c058ef8f9805daca546b', 'point.json': '37517e5f3dc66819f61f5a7bb8ace1921282415f10551d2defa5c3eb0985b570', 'point.json.lua': 'e3b0c44298fc1c149afbf4c8996fb92427ae41e4649b934ca495991b7852b855', 'prj.json': '14f1471434bc39ae6f11944fdff35eff23d14d9e65682650c694a0375f86ce9c', 'src0.lua': '481da55f95ee781931c7cefdb89dfee91854a544684f3d3b2856227ead004d9e'}


def exists(sftp, path):
    try:
        sftp.stat(path)
    except OSError as error:
        if error.errno == errno.ENOENT:
            return False
        raise
    return True


def upload(allow_create=True):
    sys.path.insert(0, str(WORKSPACE / "tools"))
    import rssh
    import paramiko

    content = {name: (PROJECT / name).read_bytes() for name in FILES}
    if {name: hashlib.sha256(data).hexdigest() for name, data in content.items()} != EXPECTED:
        raise RuntimeError("本地工程与已核对版本不一致。")
    target = REMOTE_ROOT + "/" + PROJECT_NAME
    pending = REMOTE_ROOT + "/." + PROJECT_NAME + "_" + uuid.uuid4().hex
    client = paramiko.SSHClient()
    client.set_missing_host_key_policy(paramiko.AutoAddPolicy())
    try:
        client.connect(rssh.HOST, username=rssh.USER, password=rssh.PASS,
                       timeout=8, allow_agent=False, look_for_keys=False)
        with client.open_sftp() as sftp:
            sftp.get_channel().settimeout(8)

            def verify(folder):
                for name, data in content.items():
                    with sftp.open(folder + "/" + name, "rb") as file:
                        if file.read() != data:
                            raise RuntimeError("回读不一致：" + name)

            if exists(sftp, target):
                verify(target)
                return "工程已在控制器，文件回读一致。"
            if not allow_create:
                raise RuntimeError("请先上传工程。")
            sftp.mkdir(pending)
            try:
                for name, data in content.items():
                    with sftp.open(pending + "/" + name, "wb") as file:
                        file.write(data)
                verify(pending)
                sftp.rename(pending, target)
            except Exception:
                if exists(sftp, pending):
                    for name in FILES:
                        path = pending + "/" + name
                        if exists(sftp, path):
                            sftp.remove(path)
                    sftp.rmdir(pending)
                raise
            verify(target)
            return "上传完成，控制器端 5 个文件回读一致。"
    finally:
        client.close()


def start_project():
    upload(allow_create=False)
    import rssh

    def command(connection, request):
        connection.sendall(request.encode("ascii"))
        data = b""
        while b";" not in data:
            chunk = connection.recv(4096)
            if not chunk:
                raise RuntimeError("命令口无应答，请确认 RoboDK 驱动已断开。")
            data += chunk
        return data.decode("ascii", errors="replace")

    def values(reply):
        match = re.match(r"^\s*0,\{([^}]*)\}", reply)
        if not match:
            raise RuntimeError("控制器拒绝查询：" + reply)
        return [float(value) for value in match.group(1).split(",") if value]

    with socket.create_connection((rssh.HOST, 29999), timeout=4) as connection:
        if values(command(connection, "RobotMode()")) != [5.0]:
            raise RuntimeError("控制器未处于已使能待机状态。")
        axes = values(command(connection, "GetAngle()"))
        if len(axes) != 6 or not all(abs(angle) <= 0.05 for angle in axes):
            raise RuntimeError("六轴起始角度不在零位容差内。")
        connection.sendall(("RunScript(" + PROJECT_NAME + ")").encode("ascii"))
        try:
            reply = connection.recv(4096).decode("ascii", errors="replace")
        except OSError:
            return "启动命令已发送，应答未确认。请查看控制器状态，避免重复点击。"
        if not reply:
            return "启动命令已发送，应答未确认。请查看控制器状态，避免重复点击。"
        if not re.match(r"^\s*0,", reply):
            raise RuntimeError("控制器拒绝启动：" + reply)
    return "控制器已接受启动命令。请观察零位→P3（首段直线） 的运动和到位状态。"


def run_action(action, pending, lock_start=False):
    button.configure(state="disabled")
    start_button.configure(state="disabled")
    status.set(pending)

    def worker():
        try:
            message = action()
            locked = lock_start
        except Exception as error:
            message = "操作未完成：" + str(error)
            locked = False
        try:
            window.after(0, finish, message, locked)
        except (RuntimeError, tk.TclError):
            pass

    threading.Thread(target=worker, daemon=False).start()


def finish(message, locked):
    status.set(message)
    button.configure(state="normal")
    if not locked:
        start_button.configure(state="normal")


if __name__ == "__main__":
    window = tk.Tk()
    window.title("CR5 零位→P3（首段直线） 工程上传")
    status = tk.StringVar(value="等待上传。上传与启动分开。点击启动会使实机从零位移动到 P1。")
    ttk.Label(window, text=PROJECT_NAME, padding=12).pack()
    button = ttk.Button(window, text="上传到控制器", command=lambda: run_action(upload, "正在上传并校验…"))
    button.pack(pady=5)
    start_button = ttk.Button(window, text="启动零位→P3（首段直线）（实机运动）",
                              command=lambda: run_action(start_project, "核对工程及控制器状态…", True))
    start_button.pack(pady=5)
    ttk.Label(window, textvariable=status, wraplength=480, padding=12).pack()
    window.mainloop()
